// TwinCAT 3 PLC project PLC_Tank
// ProgramVersion: 3.1.4026.27
// libraries:
//   Tc2_ControllerToolbox, * (Beckhoff Automation GmbH)
//   Tc2_ModbusSrv, * (Beckhoff Automation GmbH)
//   Tc2_Standard, * (Beckhoff Automation GmbH)
//   Tc2_System, * (Beckhoff Automation GmbH)
//   Tc3_Module, * (Beckhoff Automation GmbH)
//   VisuDialogs, * (System)
//   VisuSymbols,3.5.10.0,System
// project tree:
//   DUTs/ TAnalogConversion.TcDUT, TEngine.TcDUT, TEngineCmd.TcDUT, THeaterState.TcDUT, THeaterCmd.TcDUT, THeater.TcDUT, TPhaseHeating.TcDUT, TPhaseCmd.TcDUT, TPhaseDraining.TcDUT, TPhaseFilling.TcDUT, TPhaseMixing.TcDUT, TPhaseState.TcDUT, TValveState.TcDUT, TValveCmd.TcDUT, TEngineState.TcDUT, TTank.TcDUT, TValve.TcDUT
//   / GlobalTextList.TcGTLO, PlcTask.TcTTO, PlcTask500ms.TcTTO, VisualizationManager.TcVMO (not stored)
//   GVLs/ Global.TcGVL
//   POUs/ Draining.TcPOU, Engine_1DO.TcPOU, FB_Tank.TcPOU, Filling.TcPOU, Heater.TcPOU, Heating.TcPOU, Main_Batch.TcPOU, MB_Connector.TcPOU, Mixing.TcPOU, Test.TcPOU, Valve_2DO.TcPOU, MAIN.TcPOU
//   POUs/Misc/ EngToRaw.TcPOU, RawToEng.TcPOU
//   VISUs/ Diagnostika.TcVIS, Faze.TcVIS, Prehled.TcVIS, Zarizeni.TcVIS
// real-time tasks:
//   TASK PlcTask: cycle T#100000us, priority 20, ADS port 350
//   TASK PlcTask500ms: cycle T#500ms, priority 1, ADS port 351

CONFIGURATION PLC_Tank
    RESOURCE PLC ON TwinCAT3
        TASK PlcTask(INTERVAL := T#100000us, PRIORITY := 20);
        TASK PlcTask500ms(INTERVAL := T#500ms, PRIORITY := 1);
        PROGRAM MB_Connector WITH PlcTask : MB_Connector;
        PROGRAM Main_Batch WITH PlcTask : Main_Batch;
        PROGRAM MAIN WITH PlcTask500ms : MAIN;
    END_RESOURCE
END_CONFIGURATION

// ---- DUTs/TAnalogConversion.TcDUT
TYPE TAnalogConversion :
STRUCT
	TransducerLoLevel : UINT;
	TransducerHiLevel : UINT;
	ScaledValLoLevel : REAL;
	ScaledValHiLevel : REAL;
END_STRUCT
END_TYPE

// ---- DUTs/TEngine.TcDUT
TYPE TEngine :
STRUCT
	Cmd : TEngineCmd;
	State : TEngineState;
	Time2Start : TIME := T#5S;
	RisingEdgeTrigger : R_TRIG;
	StartupFailTimer : TON;
END_STRUCT
END_TYPE

// ---- DUTs/TEngineCmd.TcDUT
TYPE TEngineCmd :
STRUCT
		SetRT : DINT;
		AutCtrl : BOOL;
		ManCtrl : BOOL;
		TurnOnMan : BOOL;
		TurnOffMan : BOOL;
		Req2RunAutCtrl : BOOL;
		ResetSUF : BOOL;
END_STRUCT
END_TYPE

// ---- DUTs/THeaterState.TcDUT
TYPE THeaterState :
STRUCT
	EnableOut : BOOL;
	HeatingOut : REAL;
	AutCtrl : BOOL;
	ManCtrl : BOOL;
	Err 	: BOOL;
	StateInt : INT;
	GenErr : BOOL; //signalisation: error occured

	HeatingPower : REAL;
	

END_STRUCT
END_TYPE

// ---- DUTs/THeaterCmd.TcDUT
TYPE THeaterCmd :
STRUCT
	AutCtrl : BOOL;
	ManCtrl : BOOL;
	TurnOnMan : BOOL;
	TurnOffMan : BOOL;
	Req2RunAutCtrl : BOOL;
END_STRUCT
END_TYPE

// ---- DUTs/THeater.TcDUT
TYPE THeater :
STRUCT
	Cmd : THeaterCmd;
	State : THeaterState;
	
	ParamHeatingPowerManual : REAL;
	ParamHeatingSetPointAutomat : REAL;
	
	PID : FB_CTRL_PID;
	ThresholdTimer : TON;
	
END_STRUCT
END_TYPE

// ---- DUTs/TPhaseHeating.TcDUT
TYPE TPhaseHeating :
STRUCT
	Cmd : TPhaseCmd;
	State : TPhaseState;
	
	ParamReqTemp : REAL;
	
	WaterTemp : REAL;
	
	fTime : INT;
END_STRUCT
END_TYPE

// ---- DUTs/TPhaseCmd.TcDUT
TYPE TPhaseCmd :
STRUCT
	StartAut : BOOL;
	StopAut : BOOL;
	StartMan : BOOL;
	StopMan : BOOL;
	PauseMan : BOOL;
	ResumeMan : BOOL;
	ResetDone : BOOL;
	AutCtrl : BOOL;
	ManCtrl : BOOL;
END_STRUCT
END_TYPE

// ---- DUTs/TPhaseDraining.TcDUT
TYPE TPhaseDraining :
STRUCT
	Cmd : TPhaseCmd;
	State : TPhaseState;
	
	ParamDrainLevel : REAL;
	WaterLevel : REAL;
END_STRUCT
END_TYPE

// ---- DUTs/TPhaseFilling.TcDUT
TYPE TPhaseFilling :
STRUCT
	Cmd : TPhaseCmd;
	State : TPhaseState;
	
	ParamFillLevel : REAL;
	WaterLevel : REAL;
END_STRUCT
END_TYPE

// ---- DUTs/TPhaseMixing.TcDUT
TYPE TPhaseMixing :
STRUCT
	Cmd : TPhaseCmd;
	State : TPhaseState;
	
	ParamTimeSec : INT;
	
	ElapsedTimeSec : INT;
END_STRUCT
END_TYPE

// ---- DUTs/TPhaseState.TcDUT
TYPE TPhaseState :
STRUCT
	Running : BOOL;
	Idle : BOOL;
	Paused : BOOL;
	Done : BOOL;
	AutCtrl : BOOL;
	ManCtrl : BOOL;
	Stateint : INT;
END_STRUCT
END_TYPE

// ---- DUTs/TValveState.TcDUT
TYPE TValveState :
STRUCT
		Open : BOOL;
		Closed : BOOL;
		OpenOut : BOOL;
		CloseOut : BOOL;
		Err : BOOL;
		StartupFail : BOOL;
		AutCtrl : BOOL;
		ManCtrl : BOOL;
		MayRun : BOOL;
		MayAutoRun : BOOL; //device is working in automatic regime
		GenErr : BOOL; //signalisation: error occured
		StColor : INT; //valve state: Open(0), Closed(1), OpenAndErr(2), ClosedAndErr(3) ,NotOpenNotClosedNotErr(4), NotOpenNotClosedAndErr(5), OpenAndClosedAndErr(6), OpenAndClosedNotErr(7)

END_STRUCT
END_TYPE

// ---- DUTs/TValveCmd.TcDUT
TYPE TValveCmd :
STRUCT
		AutCtrl : BOOL;
		ManCtrl : BOOL;
		OpenMan : BOOL;
		StopMan : BOOL;
		CloseMan : BOOL;
		Req2OpenAut : BOOL;
		Req2CloseAut : BOOL;
		ResetSUF : BOOL;
END_STRUCT
END_TYPE

// ---- DUTs/TEngineState.TcDUT
TYPE TEngineState :
STRUCT
		RT : DINT;
		Run : BOOL;
		RunOut : BOOL;
		Err : BOOL;
		StartUpFail : BOOL;
		AutCtrl : BOOL;
		ManCtrl : BOOL;
		MayRun : BOOL;
		MayAutoRun : BOOL;
		GenErr : BOOL;
		StateInt : INT;
		
		StartupFailTime : INT;
END_STRUCT
END_TYPE

// ---- DUTs/TTank.TcDUT
TYPE TTank :
STRUCT
	Mixer : TEngine;
	ValveFilling : TValve;
	ValveDraining : TValve;
	Heater : THeater;
	
	Filling : TPhaseFilling;
	Draining : TPhaseDraining;
	Mixing : TPhaseMixing;
	Heating : TPhaseHeating;
	
	GlobalError : BOOL;

END_STRUCT
END_TYPE

// ---- DUTs/TValve.TcDUT
TYPE TValve :
STRUCT
	Cmd : TValveCmd;
	State : TValveState;
	Time2Open : TIME := T#12S;
	
	OpenFailTimer : TON;
	CloseFailTimer : TON;
	
END_STRUCT
END_TYPE

// ---- GVLs/Global.TcGVL
{attribute 'qualified_only'}
VAR_GLOBAL
	Tank1 : TTank;
	

	secImp : BOOL;
	
	diMixerRun : BOOL;
	diMixerError : BOOL;
	diValveFillOpen : BOOL;
	diValveFillClose : BOOL;
	diValveFillError : BOOL;
	diValveDrainOpen : BOOL;
	diValveDrainClose : BOOL;
	diValveDrainError : BOOL;
	
	aiWaterLevel : WORD;
	aiWaterTemp : WORD;
	
	doMixerStart : BOOL;
	doValveFillOpen : BOOL;
	doValveFillClose : BOOL;
	doValveDrainOpen : BOOL;
	doValveDrainClose : BOOL;
	doHeatingEnable : BOOL;
	
	aoReqPowerOfHeating : WORD;

END_VAR

VAR_GLOBAL CONSTANT
	Running : INT := 0;
	Stop : INT := 1;
	RunningAndError : INT := 2;
	Err : INT := 3;

	PhIdle : INT := 0;
	PhRunning : INT := 1;
	PhPause : INT := 2;
	
    Open : INT := 0;
	Closed : INT := 1;
	OpenAndErr : INT := 2;
	ClosedAndErr : INT := 3;
	NotOpenNotClosedNotErr : INT := 4;
	NotOpenNotClosedAndErr : INT := 5;
	OpenAndClosedAndErr : INT := 6;
	OpenAndClosedNotErr : INT := 7;
END_VAR

// ---- POUs/MB_Connector.TcPOU
PROGRAM MB_Connector
VAR
	
	mb_ipaddr   : STRING(15) := '127.0.0.1';
	mb_port		: UINT := 504;
	mb_unitid	: BYTE := 1;
	
	fbReadRegs		: FB_MBReadInputRegs;
	mb_regs    		: ARRAY [0..4] OF WORD;
	mb_regs_error	: BOOL;
	mb_regs_busy	: BOOL;
	mb_regs_execute : BOOL;
	mb_regs_errid	: UDINT;
	
	fbReadInps	: FB_MBReadInputs;
	mb_inps			: ARRAY [0..4] OF BYTE;
	mb_inps_error	: BOOL;
	mb_inps_busy	: BOOL;
	mb_inps_execute : BOOL;
	mb_inps_errid	: UDINT;
	
	fbWriteRegs		: FB_MBWriteRegs;
	mbw_regs    	: ARRAY [0..4] OF WORD;
	mbw_regs_error	: BOOL;
	mbw_regs_busy	: BOOL;
	mbw_regs_execute: BOOL;
	mbw_regs_errid	: UDINT;
	
	fbWriteCoils	: FB_MBWriteCoils;
	mbw_coils		: ARRAY [0..4] OF BYTE;
	mbw_coils_error	: BOOL;
	mbw_coils_busy	: BOOL;
	mbw_coils_execute: BOOL;
	mbw_coils_errid	: UDINT;
	
END_VAR

fbReadRegs.sIPAddr := mb_ipaddr;
fbReadRegs.nTCPPort := mb_port;
fbReadRegs.nQuantity := 4;
fbReadRegs.nMBAddr := 0;
fbReadRegs.cbLength := SIZEOF(mb_regs);
fbReadRegs.pDestAddr := ADR(mb_regs);
fbReadRegs.nUnitID := mb_unitid;
fbReadRegs.tTimeout := T#5S;
IF (mb_regs_busy = FALSE) THEN
	mb_regs_execute := TRUE;
ELSE
	mb_regs_execute := FALSE;
END_IF
fbReadRegs(bExecute := mb_regs_execute, 
		   bBusy => mb_regs_busy, bError => mb_regs_error, 
		   nErrId => mb_regs_errid);



fbReadInps.sIPAddr := mb_ipaddr;
fbReadInps.nTCPPort := mb_port;
fbReadInps.nQuantity := 32;
fbReadInps.nMBAddr := 0;
fbReadInps.cbLength := SIZEOF(mb_inps);
fbReadInps.pDestAddr := ADR(mb_inps);
fbReadInps.nUnitID := mb_unitid;
fbReadInps.tTimeout := T#5S;
IF (mb_inps_busy = FALSE) THEN
	mb_inps_execute := TRUE;
ELSE
	mb_inps_execute := FALSE;
END_IF
fbReadInps(bExecute := mb_inps_execute, 
	bBusy => mb_inps_busy, bError => mb_inps_error, nErrId => mb_inps_errid);

Global.diValveFillOpen := mb_inps[0].0;
Global.diValveFillClose := mb_inps[0].1;
Global.diValveFillError := mb_inps[0].2;
Global.diValveDrainOpen := mb_inps[0].3;
Global.diValveDrainClose := mb_inps[0].4;
Global.diValveDrainError := mb_inps[0].5;
Global.diMixerRun := mb_inps[0].6;
Global.diMixerError := mb_inps[0].7;

Global.aiWaterLevel := mb_regs[0];
Global.aiWaterTemp := mb_regs[2];







fbWriteRegs.sIPAddr := mb_ipaddr;
fbWriteRegs.nTCPPort := mb_port;
fbWriteRegs.nQuantity := 4;
fbWriteRegs.nMBAddr := 0;
fbWriteRegs.cbLength := SIZEOF(mbw_regs);
fbWriteRegs.pSrcAddr := ADR(mbw_regs);
fbWriteRegs.nUnitID := mb_unitid;
fbWriteRegs.tTimeout := T#5S;
IF (mbw_regs_busy = FALSE) THEN
	mbw_regs_execute := TRUE;
ELSE
	mbw_regs_execute := FALSE;
END_IF
fbWriteRegs(bExecute := mbw_regs_execute, 
		   bBusy => mbw_regs_busy, bError => mbw_regs_error, 
		   nErrId => mbw_regs_errid);



fbWriteCoils.sIPAddr := mb_ipaddr;
fbWriteCoils.nTCPPort := mb_port;
fbWriteCoils.nQuantity := 32;
fbWriteCoils.nMBAddr := 0;
fbWriteCoils.cbLength := SIZEOF(mbw_coils);
fbWriteCoils.pSrcAddr := ADR(mbw_coils);
fbWriteCoils.nUnitID := mb_unitid;
fbWriteCoils.tTimeout := T#5S;
IF (mbw_coils_busy = FALSE) THEN
	mbw_coils_execute := TRUE;
ELSE
	mbw_coils_execute := FALSE;
END_IF
fbWriteCoils(bExecute := mbw_coils_execute, 
	bBusy => mbw_coils_busy, bError => mbw_coils_error, nErrId => mbw_coils_errid);

mbw_coils[0].0 := Global.doValveFillOpen;
mbw_coils[0].1 := Global.doValveFillClose;
mbw_coils[0].2 := Global.doValveDrainOpen;
mbw_coils[0].3 := Global.doValveDrainClose;
mbw_coils[0].4 := Global.doMixerStart;
mbw_coils[0].5 := Global.doHeatingEnable;

mbw_regs[0] := Global.aoReqPowerOfHeating;

END_PROGRAM

// ---- POUs/Main_Batch.TcPOU
PROGRAM Main_Batch
VAR
	FB_Tank_1 : FB_Tank;
END_VAR

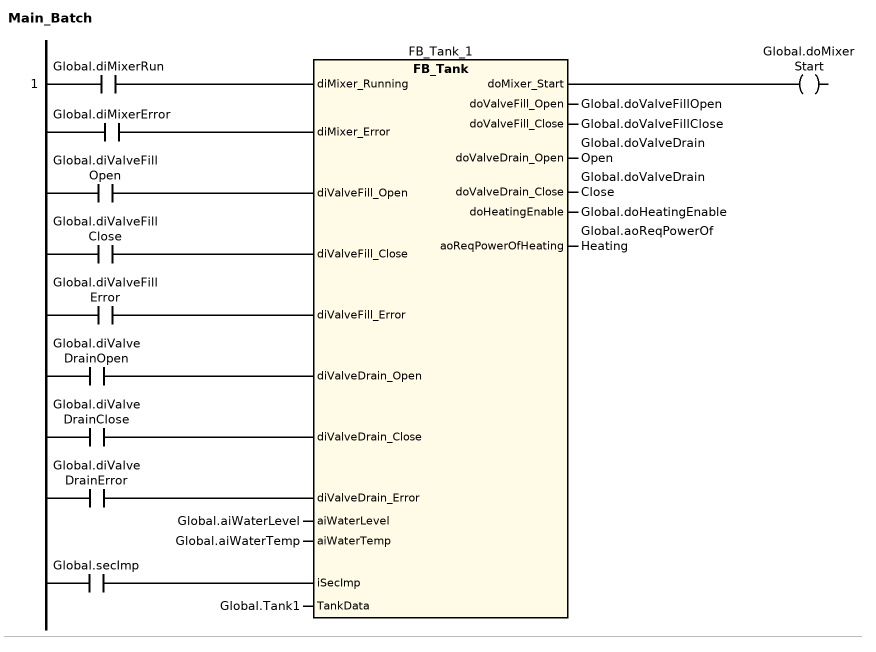
// NETWORK 1
FB_Tank_1(
    diMixer_Running := Global.diMixerRun,
    diMixer_Error := Global.diMixerError,
    diValveFill_Open := Global.diValveFillOpen,
    diValveFill_Close := Global.diValveFillClose,
    diValveFill_Error := Global.diValveFillError,
    diValveDrain_Open := Global.diValveDrainOpen,
    diValveDrain_Close := Global.diValveDrainClose,
    diValveDrain_Error := Global.diValveDrainError,
    aiWaterLevel := Global.aiWaterLevel,
    aiWaterTemp := Global.aiWaterTemp,
    iSecImp := Global.secImp,
    TankData := Global.Tank1,
    doValveFill_Open => Global.doValveFillOpen,
    doValveFill_Close => Global.doValveFillClose,
    doValveDrain_Open => Global.doValveDrainOpen,
    doValveDrain_Close => Global.doValveDrainClose,
    doHeatingEnable => Global.doHeatingEnable,
    aoReqPowerOfHeating => Global.aoReqPowerOfHeating); // FB_Tank
Global.doMixerStart := FB_Tank_1.doMixer_Start;

END_PROGRAM

// ---- POUs/FB_Tank.TcPOU
FUNCTION_BLOCK FB_Tank
VAR_INPUT
	diMixer_Running : BOOL;
	diMixer_Error : BOOL;
	diValveFill_Open : BOOL;
	diValveFill_Close : BOOL;
	diValveFill_Error : BOOL;
	diValveDrain_Open : BOOL;
	diValveDrain_Close : BOOL;
	diValveDrain_Error : BOOL;
	aiWaterLevel : WORD;
	aiWaterTemp : WORD;
	iSecImp : BOOL; //Požaduje se vstup s periodou 1 sekunda a libovolnou střídou
END_VAR

VAR_OUTPUT
	doMixer_Start : BOOL;
	doValveFill_Open : BOOL;
	doValveFill_Close : BOOL;
	doValveDrain_Open : BOOL;
	doValveDrain_Close : BOOL;
	doHeatingEnable : BOOL;
	aoReqPowerOfHeating : WORD;
END_VAR

VAR_IN_OUT
	TankData : TTank;
END_VAR

VAR
	//Konfigurace přepočtu rozsahu převodníků
	WaterTemp : TAnalogConversion := (TransducerLoLevel := 0, TransducerHiLevel := 27648, ScaledValLoLevel := 0, ScaledValHiLevel := 100);
	WaterLevel : TAnalogConversion := (TransducerLoLevel := 0, TransducerHiLevel := 27648, ScaledValLoLevel := 0, ScaledValHiLevel := 2);
	ReqOutputPower : TAnalogConversion := (ScaledValLoLevel := 0, ScaledValHiLevel := 100, TransducerLoLevel := 0, TransducerHiLevel := 27648);

	//Instance zanořených funkčních bloků
	ValveDrainCm : Valve_2DO;
	ValveFillCm : Valve_2DO;
	MixerCm : Engine_1DO;
	HeaterCm : Heater;
	FillingPhase : Filling;
	MixingPhase : Mixing;
	DrainingPhase : Draining;
	HeatingPhase : Heating;
	TON1: TON;
	RawToEng_1: RawToEng;
	RawToEng_2: RawToEng;
	EngToRaw_1: EngToRaw;
END_VAR

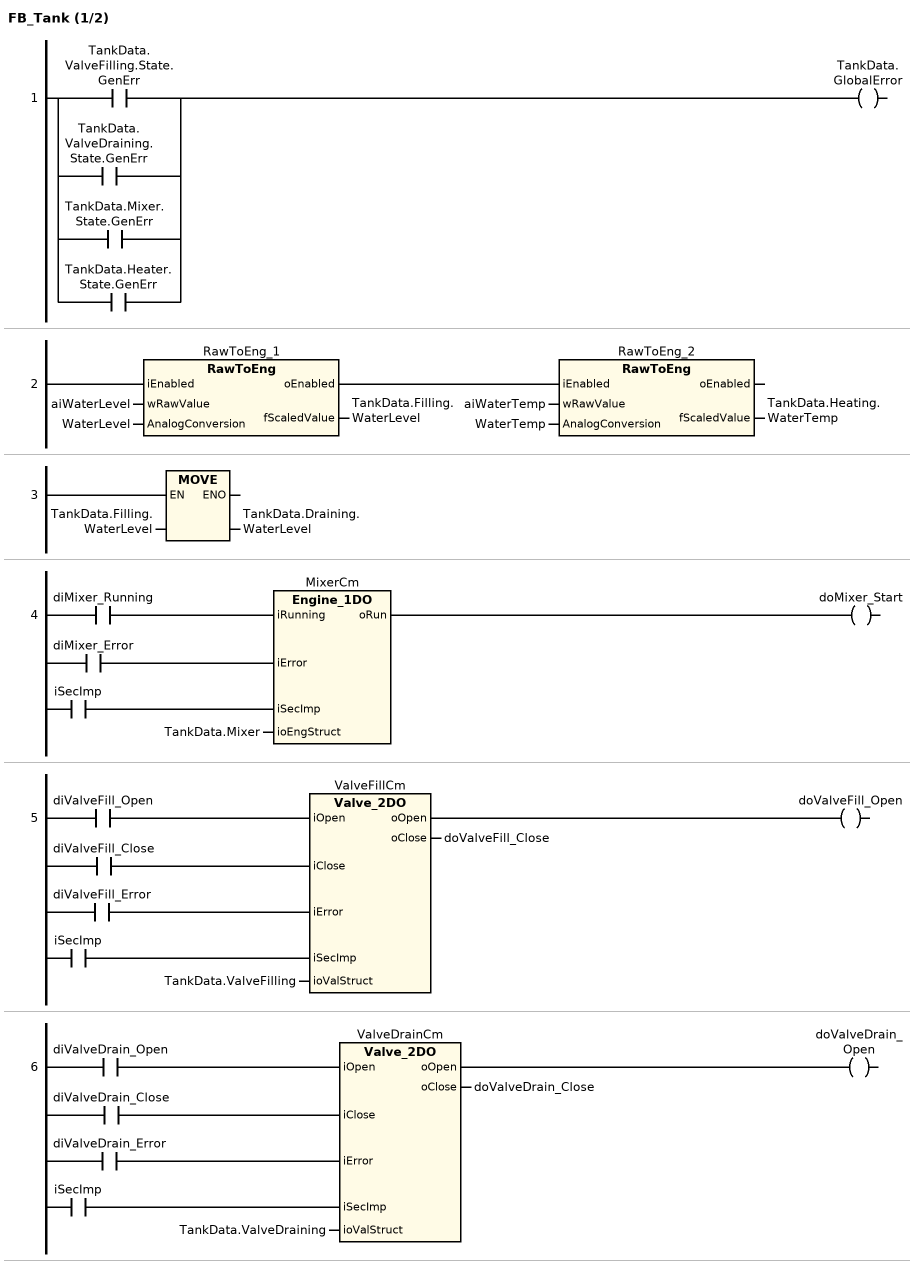
// NETWORK 1
TankData.GlobalError := TankData.ValveFilling.State.GenErr OR TankData.ValveDraining.State.GenErr OR TankData.Mixer.State.GenErr OR TankData.Heater.State.GenErr;

// NETWORK 2
RawToEng_1(
    iEnabled := TRUE,
    wRawValue := aiWaterLevel,
    AnalogConversion := WaterLevel,
    fScaledValue => TankData.Filling.WaterLevel); // RawToEng
RawToEng_2(
    iEnabled := RawToEng_1.oEnabled,
    wRawValue := aiWaterTemp,
    AnalogConversion := WaterTemp,
    fScaledValue => TankData.Heating.WaterTemp); // RawToEng

// NETWORK 3
TankData.Draining.WaterLevel := TankData.Filling.WaterLevel;

// NETWORK 4
MixerCm(
    iRunning := diMixer_Running,
    iError := diMixer_Error,
    iSecImp := iSecImp,
    ioEngStruct := TankData.Mixer); // Engine_1DO
doMixer_Start := MixerCm.oRun;

// NETWORK 5
ValveFillCm(
    iOpen := diValveFill_Open,
    iClose := diValveFill_Close,
    iError := diValveFill_Error,
    iSecImp := iSecImp,
    ioValStruct := TankData.ValveFilling,
    oClose => doValveFill_Close); // Valve_2DO
doValveFill_Open := ValveFillCm.oOpen;

// NETWORK 6
ValveDrainCm(
    iOpen := diValveDrain_Open,
    iClose := diValveDrain_Close,
    iError := diValveDrain_Error,
    iSecImp := iSecImp,
    ioValStruct := TankData.ValveDraining,
    oClose => doValveDrain_Close); // Valve_2DO
doValveDrain_Open := ValveDrainCm.oOpen;

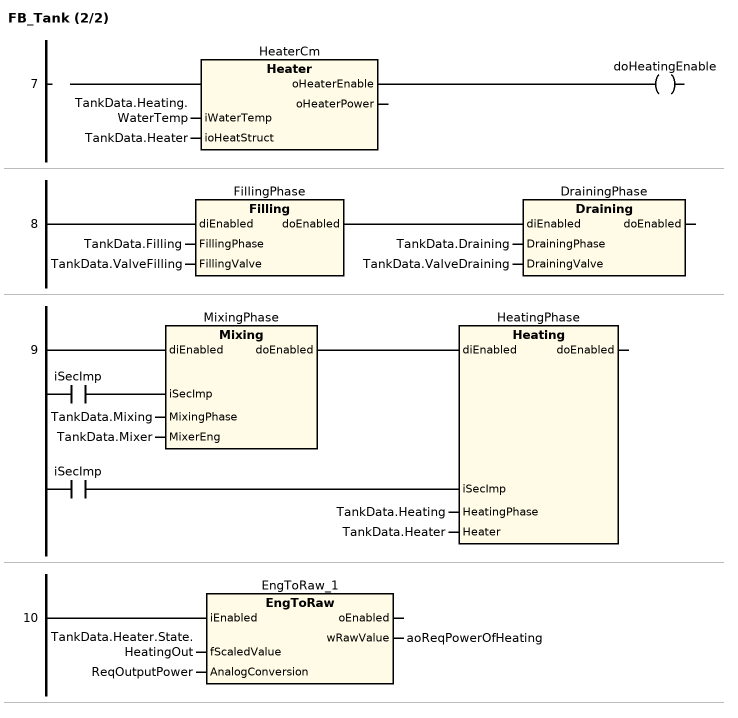
// NETWORK 7
HeaterCm(iWaterTemp := TankData.Heating.WaterTemp, ioHeatStruct := TankData.Heater); // Heater
doHeatingEnable := HeaterCm.oHeaterEnable;

// NETWORK 8
FillingPhase(diEnabled := TRUE, FillingPhase := TankData.Filling, FillingValve := TankData.ValveFilling); // Filling
DrainingPhase(
    diEnabled := FillingPhase.doEnabled,
    DrainingPhase := TankData.Draining,
    DrainingValve := TankData.ValveDraining); // Draining

// NETWORK 9
MixingPhase(
    diEnabled := TRUE,
    iSecImp := iSecImp,
    MixingPhase := TankData.Mixing,
    MixerEng := TankData.Mixer); // Mixing
HeatingPhase(
    diEnabled := MixingPhase.doEnabled,
    iSecImp := iSecImp,
    HeatingPhase := TankData.Heating,
    Heater := TankData.Heater); // Heating

// NETWORK 10
EngToRaw_1(
    iEnabled := TRUE,
    fScaledValue := TankData.Heater.State.HeatingOut,
    AnalogConversion := ReqOutputPower,
    wRawValue => aoReqPowerOfHeating); // EngToRaw

END_FUNCTION_BLOCK

// ---- POUs/Valve_2DO.TcPOU
FUNCTION_BLOCK Valve_2DO
VAR_INPUT
	iOpen : BOOL;
	iClose : BOOL;
	iError : BOOL;
	iSecImp : BOOL;
END_VAR
VAR_OUTPUT
	oOpen : BOOL;
	oClose : BOOL;
END_VAR

VAR_IN_OUT
	ioValStruct	 : TValve;
END_VAR

VAR
	tempOpenStartupFail : BOOL;
	tempCloseStartupFail: BOOL;
END_VAR

{region "OpenState"}
    // set real state of valve input into valve structure - input of valve can be taken from limit sensor...
    ioValStruct.State.Open := iOpen;
    ioValStruct.State.Closed := iClose;
{endregion}

	 
{region "REGION Aut/Man"}
    // switching state of engine - automatic or manual control (default state is manual)
  	IF ioValStruct.Cmd.ManCtrl THEN
      	ioValStruct.State.ManCtrl := TRUE;
		ioValStruct.State.AutCtrl := FALSE;
	ELSIF ioValStruct.Cmd.AutCtrl THEN
        ioValStruct.State.ManCtrl := FALSE;
		ioValStruct.State.AutCtrl := TRUE; 
    END_IF;
		 
	IF (NOT ioValStruct.State.AutCtrl AND NOT ioValStruct.State.ManCtrl) THEN
		ioValStruct.State.ManCtrl := TRUE;
	END_IF

	ioValStruct.Cmd.ManCtrl := FALSE;
	ioValStruct.Cmd.AutCtrl := FALSE;
{endregion}
	 
{region "MayRun / MayAutoRun"}
    // setting auxilary signals (may run, may auto run) - MR AND NOT MAR - engine may be started in manual mode, MAR - engine may be started in automatic mode
    ioValStruct.State.MayRun := (ioValStruct.State.ManCtrl AND NOT(ioValStruct.State.GenErr));
	ioValStruct.State.MayAutoRun := (ioValStruct.State.AutCtrl AND NOT(ioValStruct.State.GenErr));
{endregion}
	 
{region "ManCtrl"}
	// processing manual actions - if command is processed, it is sets to FALSE even if can't be processed
    // Valve commands are open, close and stop - valve can be stopped intermediate position
	 IF ioValStruct.State.ManCtrl AND ioValStruct.State.MayRun THEN
        IF ioValStruct.Cmd.OpenMan THEN
            ioValStruct.State.CloseOut := FALSE;
            ioValStruct.State.OpenOut := TRUE;
        END_IF;
        
        IF ioValStruct.Cmd.CloseMan THEN
            ioValStruct.State.OpenOut := FALSE;
            ioValStruct.State.CloseOut := TRUE;
        END_IF;
        
        IF ioValStruct.Cmd.StopMan THEN
            ioValStruct.State.OpenOut := FALSE;
            ioValStruct.State.CloseOut := FALSE;
        END_IF;
    END_IF;
    
    ioValStruct.Cmd.OpenMan := FALSE;
    ioValStruct.Cmd.CloseMan := FALSE;
    ioValStruct.Cmd.StopMan := FALSE;
{endregion}
	 
{region "AutCtrl"}
	 //if request to run in automatic mode -> set outputs to right states if MAR
    //AutoRequest shouldn't be reseted to false state
    //if request to open and request to close are setted to 1 simultaneously - outputs should be 0.
    IF ioValStruct.State.AutCtrl AND ioValStruct.State.MayAutoRun THEN
        IF ioValStruct.Cmd.Req2CloseAut AND (NOT ioValStruct.Cmd.Req2OpenAut) THEN
            ioValStruct.State.OpenOut := FALSE;
            ioValStruct.State.CloseOut := TRUE;
        END_IF;
        
        IF (NOT ioValStruct.Cmd.Req2CloseAut) AND ioValStruct.Cmd.Req2OpenAut THEN
            ioValStruct.State.CloseOut := FALSE;
            ioValStruct.State.OpenOut := TRUE;
        END_IF;
        
        IF (NOT ioValStruct.Cmd.Req2CloseAut) AND (NOT ioValStruct.Cmd.Req2OpenAut) THEN
            ioValStruct.State.CloseOut := FALSE;
            ioValStruct.State.OpenOut := FALSE;
        END_IF;
        
    END_IF;
{endregion}
	 
{region "Error states"}
 // definition of error states 
    // error - input from digital input of plc - fyzical state of valve
    // calculating start up fail - if output is sets to open or close, it's expected feedback from limit sensor in defined time, if feedback doesn't show in this time, it should be start up fail error
    // merge of these two error is general error
    // error is both inputs (open and closed) true state
    ioValStruct.OpenFailTimer(IN := ioValStruct.State.OpenOut AND NOT ioValStruct.State.CloseOut AND NOT ioValStruct.State.Open, PT := ioValStruct.Time2Open);
	tempOpenStartupFail := ioValStruct.OpenFailTimer.Q;

    ioValStruct.CloseFailTimer(IN := ioValStruct.State.CloseOut AND NOT ioValStruct.State.OpenOut AND NOT ioValStruct.State.Closed, PT := ioValStruct.Time2Open);
	tempCloseStartupFail := ioValStruct.CloseFailTimer.Q;
    
   
    IF tempOpenStartupFail OR tempCloseStartupFail THEN
        ioValStruct.State.StartUpFail := TRUE;
    END_IF;
    
    IF iError THEN
        ioValStruct.State.Err := TRUE;
    END_IF;
    
    ioValStruct.State.GenErr := ioValStruct.State.StartUpFail OR iError;
    
    // start up fail can be reseted by operator, command resetSUF, resets SUF and engine should be started again
    IF ioValStruct.Cmd.ResetSUF THEN
        ioValStruct.State.StartUpFail := FALSE;
        ioValStruct.Cmd.ResetSUF := FALSE;
    END_IF;
    
    // if error state exists outputs should be in stop state
    IF ioValStruct.State.GenErr THEN
        ioValStruct.State.OpenOut := FALSE;
        ioValStruct.State.CloseOut := FALSE;
    END_IF;
{endregion}
	 	 
oOpen := ioValStruct.State.OpenOut;
oClose := ioValStruct.State.CloseOut;

{region "StatusInt"}
    //write combination of states into int value for visualization (valve - combination of open, close state and error)
    IF ioValStruct.State.Open AND NOT ioValStruct.State.Closed AND NOT ioValStruct.State.GenErr THEN
        ioValStruct.State.StColor := Global.Open;
    ELSIF NOT ioValStruct.State.Open AND ioValStruct.State.Closed AND NOT ioValStruct.State.GenErr THEN
        ioValStruct.State.StColor := Global.Closed;
    ELSIF ioValStruct.State.Open AND NOT ioValStruct.State.Closed AND ioValStruct.State.GenErr THEN
        ioValStruct.State.StColor := Global.OpenAndErr;
    ELSIF NOT ioValStruct.State.Open AND ioValStruct.State.Closed AND ioValStruct.State.GenErr THEN
        ioValStruct.State.StColor := Global.ClosedAndErr;
    ELSIF NOT ioValStruct.State.Open AND NOT ioValStruct.State.Closed AND NOT ioValStruct.State.GenErr THEN
        ioValStruct.State.StColor := Global.NotOpenNotClosedNotErr;
    ELSIF NOT ioValStruct.State.Open AND NOT ioValStruct.State.Closed AND ioValStruct.State.GenErr THEN
        ioValStruct.State.StColor := Global.NotOpenNotClosedAndErr;
    ELSIF ioValStruct.State.Open AND ioValStruct.State.Closed AND ioValStruct.State.GenErr THEN
        ioValStruct.State.StColor := Global.OpenAndClosedAndErr;
    ELSIF ioValStruct.State.Open AND ioValStruct.State.Closed AND NOT ioValStruct.State.GenErr THEN
        ioValStruct.State.StColor := Global.OpenAndClosedNotErr;
    END_IF;
{endregion}

END_FUNCTION_BLOCK

// ---- POUs/Engine_1DO.TcPOU
FUNCTION_BLOCK Engine_1DO
VAR_INPUT
	iRunning : BOOL;
	iError : BOOL;
	iSecImp : BOOL;
END_VAR
VAR_OUTPUT
	oRun : BOOL;
END_VAR
VAR_IN_OUT
	ioEngStruct : TEngine;
END_VAR
VAR
	secImpEdge: BOOL;
	tempStartupFail: BOOL;
END_VAR

{region "RunState"}
    // set real state of engine run into engine structure
  ioEngStruct.State.Run := iRunning;
{endregion}

{region "Running time"} 
    // counting running time of engine - (motoseconds in real situation it should be moto hours)
    // detection rising edge of input secimp - should be conected 1Hz internal clock from PLC
	IF ioEngStruct.State.Run THEN
		IF iSecImp AND NOT secImpEdge THEN
			secImpEdge := TRUE;
			ioEngStruct.State.RT := ioEngStruct.State.RT + 1;
		ELSIF NOT iSecImp THEN
			secImpEdge := FALSE; 
		END_IF
	END_IF 
	
	IF ioEngStruct.Cmd.SetRT >= 0 THEN
		ioEngStruct.State.RT := ioEngStruct.Cmd.SetRT;
		ioEngStruct.Cmd.SetRT := -1;
	END_IF
{endregion}
	 
 
{region "Manual/Automat"}
	// switching state of engine - automatic or manual control (default state is manual)
	IF ioEngStruct.Cmd.ManCtrl THEN
      	ioEngStruct.State.ManCtrl := TRUE;
		ioEngStruct.State.AutCtrl := FALSE;
	ELSIF ioEngStruct.Cmd.AutCtrl THEN
        ioEngStruct.State.ManCtrl := FALSE;
		ioEngStruct.State.AutCtrl := TRUE; 
    END_IF;
		 
	IF (NOT ioEngStruct.State.AutCtrl AND NOT ioEngStruct.State.ManCtrl) THEN
		ioEngStruct.State.ManCtrl := TRUE;
	END_IF

	ioEngStruct.Cmd.ManCtrl := FALSE;
	ioEngStruct.Cmd.AutCtrl := FALSE;
{endregion}
	 
{region "MayRun / MayAutoRun"}
	// setting auxilary signals (may run, may auto run) - MR AND NOT MAR - eng should be started in manual mode,
    // MAR - should be started in automatic mode
    ioEngStruct.State.MayRun := (ioEngStruct.State.ManCtrl AND NOT(ioEngStruct.State.GenErr));
	ioEngStruct.State.MayAutoRun := (ioEngStruct.State.AutCtrl AND NOT(ioEngStruct.State.GenErr));  
{endregion}
	 
{region "ManCtrl"}
	// processing manual actions - if command is processed, it is set to FALSE even if can't be processed
    // Engine commands are turn off (stop) and turn on (start)
	IF ioEngStruct.State.ManCtrl AND ioEngStruct.State.MayRun THEN
		IF ioEngStruct.Cmd.TurnOnMan THEN
			ioEngStruct.State.RunOut := TRUE;
		ELSIF ioEngStruct.Cmd.TurnOffMan THEN
			ioEngStruct.State.RunOut := FALSE;
		END_IF
    END_IF;
	ioEngStruct.Cmd.TurnOnMan := FALSE;
	ioEngStruct.Cmd.TurnOffMan := FALSE;
{endregion}
	 
{region "AutCtrl"}
	//if request to run in automatic mode set outputs to right states if MAR
    //AutoRequest shouldn't be reseted to false state
    IF ioEngStruct.State.AutCtrl AND ioEngStruct.State.MayAutoRun THEN
		IF ioEngStruct.Cmd.Req2RunAutCtrl THEN
			ioEngStruct.State.RunOut := TRUE;
		ELSIF NOT ioEngStruct.Cmd.Req2RunAutCtrl THEN
			ioEngStruct.State.RunOut := FALSE;
		END_IF
    END_IF;
{endregion}
	 
{region "Error states"}
	// definition of error states 
	// error - input from digital input of plc - fyzical state of engine 
	// calculating start up fail - if output is sets to start engine, it's expected feedback from running signal in defined time, if feedback doesn't show in this time, it should be start up fail error
	// merge of these two error is general error
	ioEngStruct.StartupFailTimer(IN := ioEngStruct.State.RunOut AND NOT iRunning, PT := ioEngStruct.Time2Start);
    IF ioEngStruct.StartupFailTimer.Q THEN
        ioEngStruct.State.StartUpFail := TRUE;
    END_IF;

    ioEngStruct.State.Err := iError;
    ioEngStruct.State.GenErr := ioEngStruct.State.StartUpFail OR iError;

    IF ioEngStruct.Cmd.ResetSUF THEN
        ioEngStruct.State.StartUpFail := FALSE;
        ioEngStruct.Cmd.ResetSUF := FALSE;
    END_IF;

    IF ioEngStruct.State.GenErr THEN
        ioEngStruct.State.RunOut := FALSE;
    END_IF;
{endregion}
	 
oRun := ioEngStruct.State.RunOut;

{region "StatusInt"}
 IF NOT ioEngStruct.State.GenErr THEN
        IF ioEngStruct.State.Run THEN
            ioEngStruct.State.StateInt := Global.Running;
        ELSE
            ioEngStruct.State.StateInt := Global.Stop;
        END_IF;
    ELSE
        IF ioEngStruct.State.Run THEN
            ioEngStruct.State.StateInt := Global.RunningAndError;
        ELSE
            ioEngStruct.State.StateInt := Global.Err;
        END_IF;
    END_IF; 
{endregion}

END_FUNCTION_BLOCK

// ---- POUs/Heater.TcPOU
FUNCTION_BLOCK Heater
VAR_INPUT
	iWaterTemp : REAL;
END_VAR
VAR_OUTPUT
	oHeaterEnable : BOOL;
	oHeaterPower : REAL;
END_VAR
VAR_IN_OUT
	ioHeatStruct : THeater;
END_VAR
VAR
	pidParameters : ST_CTRL_PID_PARAMS;
	pidMode : E_CTRL_MODE;      // ACTIVE when heater is enabled, RESET otherwise
END_VAR

pidParameters.fKp := 1.196; //P
pidParameters.tTn := T#75.798S; //I
pidParameters.tTv := T#0S; //D
pidParameters.tCtrlCycleTime := T#200MS;
pidParameters.tTaskCycleTime := T#100MS;
pidParameters.fOutMaxLimit := 100;
pidParameters.fOutMinLimit := 0;
pidParameters.bDInTheFeedbackPath := FALSE;
pidParameters.bPInTheFeedbackPath := FALSE;
pidParameters.bARWOnIPartOnly := FALSE;
pidParameters.tTd := T#100MS; 


// PID runs only when heater is enabled - otherwise it is held in reset,
// so the integral part doesn't wind up while heating is off (no overshoot after start)
IF ioHeatStruct.State.EnableOut THEN
	pidMode := E_CTRL_MODE.eCTRL_MODE_ACTIVE;
ELSE
	pidMode := E_CTRL_MODE.eCTRL_MODE_RESET;
END_IF;

ioHeatStruct.PID(
	fSetpointValue := ioHeatStruct.ParamHeatingSetPointAutomat, 
	fActualValue := iWaterTemp, 
	fManSyncValue := ioHeatStruct.ParamHeatingPowerManual,
	bSync := ioHeatStruct.State.ManCtrl,
	eMode := pidMode, // automatic mode of PID component
	stParams := pidParameters);

ioHeatStruct.State.HeatingOut := ioHeatStruct.PID.fOut;

	 
{region "Manual/Automat"}
// switching state of engine - automatic or manual control (default state is manual)
	IF ioHeatStruct.Cmd.ManCtrl THEN
      	ioHeatStruct.State.ManCtrl := TRUE;
		ioHeatStruct.State.AutCtrl := FALSE;
	ELSIF ioHeatStruct.Cmd.AutCtrl THEN
        ioHeatStruct.State.ManCtrl := FALSE;
		ioHeatStruct.State.AutCtrl := TRUE; 
    END_IF;
		 
	IF (NOT ioHeatStruct.State.AutCtrl AND NOT ioHeatStruct.State.ManCtrl) THEN
		ioHeatStruct.State.ManCtrl := TRUE;
	END_IF

	ioHeatStruct.Cmd.ManCtrl := FALSE;
	ioHeatStruct.Cmd.AutCtrl := FALSE;
{endregion}
	 
 
{region "ManCtrl"}
	// processing manual actions - if command is processed, it is set to FALSE even if can't be processed
	// Heater commands are turn off (stop) and turn on (start) and power level
	IF ioHeatStruct.State.ManCtrl THEN
		IF ioHeatStruct.Cmd.TurnOnMan AND NOT ioHeatStruct.State.GenErr THEN
			ioHeatStruct.State.EnableOut := TRUE;
		ELSIF ioHeatStruct.Cmd.TurnOffMan THEN
			ioHeatStruct.State.EnableOut := FALSE;
		END_IF
    END_IF;
	ioHeatStruct.Cmd.TurnOnMan := FALSE;
	ioHeatStruct.Cmd.TurnOffMan := FALSE;
{endregion}
 
{region "AutCtrl"}
	//if request to run in automatic mode set outputs to right states if MAR
	//AutoRequest shouldn't be reseted to false state
    IF ioHeatStruct.State.AutCtrl THEN
		IF ioHeatStruct.Cmd.Req2RunAutCtrl AND NOT ioHeatStruct.State.GenErr THEN
			ioHeatStruct.State.EnableOut := TRUE;
		ELSIF NOT ioHeatStruct.Cmd.Req2RunAutCtrl THEN
			ioHeatStruct.State.EnableOut := FALSE;
		END_IF
    END_IF;
{endregion}
 
{region "Error states"}
	// if water temperature is too high, stop heating and generate error
	IF iWaterTemp > 90 THEN
		ioHeatStruct.State.EnableOut := FALSE;
		ioHeatStruct.State.GenErr := TRUE;
	ELSIF iWaterTemp < 85 THEN
		ioHeatStruct.State.GenErr := FALSE;
	END_IF
	ioHeatStruct.State.Err := ioHeatStruct.State.GenErr;
{endregion}
	 
 IF NOT ioHeatStruct.State.EnableOut THEN
    ioHeatStruct.State.HeatingOut := 0;
ELSIF ioHeatStruct.State.ManCtrl THEN
    ioHeatStruct.State.HeatingOut := ioHeatStruct.ParamHeatingPowerManual;
ELSE
    ioHeatStruct.State.HeatingOut := ioHeatStruct.PID.fOut;
END_IF;
 
oHeaterPower := ioHeatStruct.State.HeatingOut;
oHeaterEnable := ioHeatStruct.State.EnableOut;

END_FUNCTION_BLOCK

// ---- POUs/Filling.TcPOU
FUNCTION_BLOCK Filling
VAR_INPUT
	diEnabled : BOOL;
END_VAR
VAR_OUTPUT
	doEnabled : BOOL;
END_VAR
VAR_IN_OUT
	FillingPhase : TPhaseFilling;
	FillingValve : TValve;
END_VAR
VAR
END_VAR

{region "REGION Aut/Man"}
    // switching state of engine - automatic or manual control (default state is manual)
  	IF FillingPhase.Cmd.ManCtrl THEN
      	FillingPhase.State.ManCtrl := TRUE;
		FillingPhase.State.AutCtrl := FALSE;
	ELSIF FillingPhase.Cmd.AutCtrl THEN
        FillingPhase.State.ManCtrl := FALSE;
		FillingPhase.State.AutCtrl := TRUE; 
    END_IF;
		 
	IF (NOT FillingPhase.State.AutCtrl AND NOT FillingPhase.State.ManCtrl) THEN
		FillingPhase.State.ManCtrl := TRUE;
	END_IF

	FillingPhase.Cmd.ManCtrl := FALSE;
	FillingPhase.Cmd.AutCtrl := FALSE;
{endregion}

{region "ManCtrl"}
    // processing manual actions - if command is processed, it is sets to FALSE even if can't be processed
    // Phase commands are start, stop, pause and resume 
    // Start - open filling valve 
    // Stop - close filling valve
    // Pause - close filling valve
    // Resume - open filling valve
    // real states of phase are wrote into states in phase structure
    IF FillingPhase.State.ManCtrl THEN
		IF FillingPhase.State.Idle AND FillingPhase.Cmd.StartMan THEN
			FillingPhase.State.Running := TRUE;
			FillingPhase.State.Idle := FALSE;
			FillingPhase.State.Paused := FALSE;
		 	FillingPhase.State.Done := FALSE;
		ELSIF FillingPhase.Cmd.StopMan THEN
			FillingPhase.State.Running := FALSE;
			FillingPhase.State.Idle := TRUE;
			FillingPhase.State.Paused := FALSE;
		ELSIF FillingPhase.State.Running AND FillingPhase.Cmd.PauseMan THEN
			FillingPhase.State.Running := FALSE;
			FillingPhase.State.Idle := FALSE;
			FillingPhase.State.Paused := TRUE;
		ELSIF FillingPhase.State.Paused AND FillingPhase.Cmd.ResumeMan THEN
			FillingPhase.State.Running := TRUE;
			FillingPhase.State.Idle := FALSE;
			FillingPhase.State.Paused := FALSE;
			FillingPhase.State.Done := FALSE;
		END_IF
    END_IF;
	
	FillingPhase.Cmd.StartMan := FALSE;
	FillingPhase.Cmd.StopMan := FALSE;
	FillingPhase.Cmd.PauseMan := FALSE;
	FillingPhase.Cmd.ResumeMan := FALSE;
{endregion}

{region "AutCtrl"}
    // if request to run in automatic mode and phase can be run in automatic mode switch phase to running
    IF FillingPhase.State.AutCtrl THEN
		IF FillingPhase.State.Idle AND FillingPhase.Cmd.StartAut THEN
			FillingPhase.State.Running := TRUE;
			FillingPhase.State.Idle := FALSE;
		 	FillingPhase.State.Done := FALSE;
		ELSIF FillingPhase.Cmd.StopAut THEN
			FillingPhase.State.Running := FALSE;
			FillingPhase.State.Idle := TRUE;
			FillingPhase.State.Paused := FALSE;
		END_IF
    END_IF;
	
	FillingPhase.Cmd.StartAut := FALSE;
	FillingPhase.Cmd.StopAut := FALSE;
{endregion}

{region "Done"}
    //every phase should have finish condition - filling phase - if water level is above requested level
    //after that done state should be set to 1
    IF FillingPhase.State.Running AND (FillingPhase.WaterLevel >= FillingPhase.ParamFillLevel - 0.083) THEN // edit based on speed of simulation 
        FillingPhase.Cmd.StopMan := TRUE;
        FillingPhase.Cmd.StopAut := TRUE;
        FillingPhase.State.Done := TRUE;
    END_IF;

    IF FillingPhase.Cmd.ResetDone THEN
        FillingPhase.State.Done := FALSE;
        FillingPhase.Cmd.ResetDone := FALSE;
    END_IF;
{endregion}

{region "States"}
	//Command valve in cases of states
    IF FillingPhase.State.Running THEN
        FillingValve.Cmd.Req2OpenAut := TRUE;
        FillingValve.Cmd.Req2CloseAut := FALSE;
    ELSE
        FillingValve.Cmd.Req2OpenAut := FALSE;
        FillingValve.Cmd.Req2CloseAut := TRUE;
    END_IF;
{endregion}


// delault state of phase - if not any state sets state to idle
IF NOT FillingPhase.State.Idle AND NOT FillingPhase.State.Paused AND NOT FillingPhase.State.Running THEN
    FillingPhase.State.Idle := 1;
END_IF;

// write binary states into int value for visualization
IF FillingPhase.State.Idle THEN
    FillingPhase.State.Stateint := Global.PhIdle;
ELSIF FillingPhase.State.Running THEN
    FillingPhase.State.Stateint := Global.PhRunning;
ELSE
    FillingPhase.State.Stateint := Global.PhPause;
END_IF;

// Ponechte pro moznost retezeni volani bloku v LAD
doEnabled := diEnabled;

END_FUNCTION_BLOCK

// ---- POUs/Mixing.TcPOU
FUNCTION_BLOCK Mixing
VAR_INPUT
	diEnabled : BOOL;
	iSecImp : BOOL;
END_VAR
VAR_OUTPUT
	doEnabled : BOOL;
END_VAR
VAR_IN_OUT
	MixingPhase : TPhaseMixing;
	MixerEng : TEngine;
END_VAR
VAR
	rtSecImp : R_TRIG;          // rising edge of second impulse
END_VAR

{region "Aut/Man"}
    // switching state of phase - automatic or manual control (default state is manual)
    // if both commands come at once, manual has priority (safety)
    IF MixingPhase.Cmd.ManCtrl THEN
        MixingPhase.State.ManCtrl := TRUE;
        MixingPhase.State.AutCtrl := FALSE;
    ELSIF MixingPhase.Cmd.AutCtrl THEN
        MixingPhase.State.ManCtrl := FALSE;
        MixingPhase.State.AutCtrl := TRUE;
    END_IF;

    // initialization - if neither mode is active, use manual
    IF NOT MixingPhase.State.AutCtrl AND NOT MixingPhase.State.ManCtrl THEN
        MixingPhase.State.ManCtrl := TRUE;
    END_IF;

    // commands are always reset after processing
    MixingPhase.Cmd.ManCtrl := FALSE;
    MixingPhase.Cmd.AutCtrl := FALSE;
{endregion}

{region "ManCtrl"}
    // processing manual actions - if command is processed, it is set to FALSE even if can't be processed
    // Phase commands are start, stop, pause and resume
    // Start  - start mixing (elapsed time starts from 0)
    // Stop   - stop mixing
    // Pause  - stop mixing (elapsed time is kept)
    // Resume - start mixing (continues for the remaining time)
    IF MixingPhase.State.ManCtrl THEN
        IF MixingPhase.State.Idle AND MixingPhase.Cmd.StartMan THEN
            MixingPhase.State.Running := TRUE;
            MixingPhase.State.Idle := FALSE;
            MixingPhase.State.Paused := FALSE;
            MixingPhase.State.Done := FALSE;
            MixingPhase.ElapsedTimeSec := 0;
        ELSIF MixingPhase.Cmd.StopMan THEN
            MixingPhase.State.Running := FALSE;
            MixingPhase.State.Idle := TRUE;
            MixingPhase.State.Paused := FALSE;
        ELSIF MixingPhase.State.Running AND MixingPhase.Cmd.PauseMan THEN
            MixingPhase.State.Running := FALSE;
            MixingPhase.State.Idle := FALSE;
            MixingPhase.State.Paused := TRUE;
        ELSIF MixingPhase.State.Paused AND MixingPhase.Cmd.ResumeMan THEN
            MixingPhase.State.Running := TRUE;
            MixingPhase.State.Idle := FALSE;
            MixingPhase.State.Paused := FALSE;
            MixingPhase.State.Done := FALSE;
        END_IF;
    END_IF;

    MixingPhase.Cmd.StartMan := FALSE;
    MixingPhase.Cmd.StopMan := FALSE;
    MixingPhase.Cmd.PauseMan := FALSE;
    MixingPhase.Cmd.ResumeMan := FALSE;
{endregion}

{region "AutCtrl"}
    // if phase is in automatic mode, process StartAut / StopAut (from MES)
    // commands are set to FALSE after their processing
    IF MixingPhase.State.AutCtrl THEN
        IF MixingPhase.State.Idle AND MixingPhase.Cmd.StartAut THEN
            MixingPhase.State.Running := TRUE;
            MixingPhase.State.Idle := FALSE;
            MixingPhase.State.Done := FALSE;
            MixingPhase.ElapsedTimeSec := 0;
        ELSIF MixingPhase.Cmd.StopAut THEN
            MixingPhase.State.Running := FALSE;
            MixingPhase.State.Idle := TRUE;
            MixingPhase.State.Paused := FALSE;
        END_IF;
    END_IF;

    MixingPhase.Cmd.StartAut := FALSE;
    MixingPhase.Cmd.StopAut := FALSE;
{endregion}

{region "Done"}
    // every phase should have finish condition - mixing phase - elapsed running time >= requested time
    // elapsed time is counted only while running (second impulse rising edge),
    // it is kept during pause and reset only on start
    rtSecImp(CLK := iSecImp);   // must be called every cycle, otherwise edges are lost

    IF MixingPhase.State.Running AND rtSecImp.Q THEN
        MixingPhase.ElapsedTimeSec := MixingPhase.ElapsedTimeSec + 1;
    END_IF;

    // finish condition met -> stop phase (processed next cycle) and signal Done
    IF MixingPhase.State.Running AND (MixingPhase.ElapsedTimeSec >= MixingPhase.ParamTimeSec) THEN
        MixingPhase.Cmd.StopMan := TRUE;
        MixingPhase.Cmd.StopAut := TRUE;
        MixingPhase.State.Done := TRUE;
    END_IF;

    // command reset done resets done state and then resets command
    IF MixingPhase.Cmd.ResetDone THEN
        MixingPhase.State.Done := FALSE;
        MixingPhase.Cmd.ResetDone := FALSE;
    END_IF;
{endregion}

{region "States"}
    // Command mixer in cases of states
    // Running - mixer runs
    // Idle    - mixer stopped
    // Paused  - mixer stopped
    IF MixingPhase.State.Running THEN
        MixerEng.Cmd.Req2RunAutCtrl := TRUE;
    ELSE
        MixerEng.Cmd.Req2RunAutCtrl := FALSE;
    END_IF;
{endregion}

// default state of phase - if not any state sets state to idle
IF NOT MixingPhase.State.Idle AND NOT MixingPhase.State.Paused AND NOT MixingPhase.State.Running THEN
    MixingPhase.State.Idle := 1;
END_IF;

// write binary states into int value for visualization
IF MixingPhase.State.Idle THEN
    MixingPhase.State.Stateint := Global.PhIdle;
ELSIF MixingPhase.State.Running THEN
    MixingPhase.State.Stateint := Global.PhRunning;
ELSE
    MixingPhase.State.Stateint := Global.PhPause;
END_IF;

doEnabled := diEnabled;

END_FUNCTION_BLOCK

// ---- POUs/Draining.TcPOU
FUNCTION_BLOCK Draining
VAR_INPUT
	diEnabled : BOOL;
END_VAR
VAR_OUTPUT
	doEnabled : BOOL;
END_VAR
VAR_IN_OUT
	DrainingPhase : TPhaseDraining;
	DrainingValve : TValve;
END_VAR
VAR
END_VAR

{region "Aut/Man"}
    // switching state of engine - automatic or manual control (default state is manual)
  	IF DrainingPhase.Cmd.ManCtrl THEN
      	DrainingPhase.State.ManCtrl := TRUE;
		DrainingPhase.State.AutCtrl := FALSE;
	ELSIF DrainingPhase.Cmd.AutCtrl THEN
        DrainingPhase.State.ManCtrl := FALSE;
		DrainingPhase.State.AutCtrl := TRUE; 
    END_IF;
		 
	IF (NOT DrainingPhase.State.AutCtrl AND NOT DrainingPhase.State.ManCtrl) THEN
		DrainingPhase.State.ManCtrl := TRUE;
	END_IF

	DrainingPhase.Cmd.ManCtrl := FALSE;
	DrainingPhase.Cmd.AutCtrl := FALSE;
{endregion}

{region "ManCtrl"}
    // processing manual actions - if command is processed, it is sets to FALSE even if can't be processed
    // Phase commands are start, stop, pause and resume 
    // Start - open draining valve 
    // Stop - close draining valve
    // Pause - close draining valve
    // Resume - open draining valve
    // real states of phase are writed into states in phase structure
    IF DrainingPhase.State.ManCtrl THEN
		IF DrainingPhase.State.Idle AND DrainingPhase.Cmd.StartMan THEN
			DrainingPhase.State.Running := TRUE;
			DrainingPhase.State.Idle := FALSE;
			DrainingPhase.State.Paused := FALSE;
		 	DrainingPhase.State.Done := FALSE;
		ELSIF DrainingPhase.Cmd.StopMan THEN
			DrainingPhase.State.Running := FALSE;
			DrainingPhase.State.Idle := TRUE;
			DrainingPhase.State.Paused := FALSE;
		ELSIF DrainingPhase.State.Running AND DrainingPhase.Cmd.PauseMan THEN
			DrainingPhase.State.Running := FALSE;
			DrainingPhase.State.Idle := FALSE;
			DrainingPhase.State.Paused := TRUE;
		ELSIF DrainingPhase.State.Paused AND DrainingPhase.Cmd.ResumeMan THEN
			DrainingPhase.State.Running := TRUE;
			DrainingPhase.State.Idle := FALSE;
			DrainingPhase.State.Paused := FALSE;
			DrainingPhase.State.Done := FALSE;
		END_IF
    END_IF;
	
	DrainingPhase.Cmd.StartMan := FALSE;
	DrainingPhase.Cmd.StopMan := FALSE;
	DrainingPhase.Cmd.PauseMan := FALSE;
	DrainingPhase.Cmd.ResumeMan := FALSE;
{endregion}

{region "AutCtrl"}
    //if request to run in automatic mode -> set auto request to open of filling valve to 1 and close to 0, if not open 0 close 1
    // commands should be sets to false after their processing
    IF DrainingPhase.State.AutCtrl THEN
		IF DrainingPhase.State.Idle AND DrainingPhase.Cmd.StartAut THEN
			DrainingPhase.State.Running := TRUE;
			DrainingPhase.State.Idle := FALSE;
		 	DrainingPhase.State.Done := FALSE;
		ELSIF DrainingPhase.Cmd.StopAut THEN
			DrainingPhase.State.Running := FALSE;
			DrainingPhase.State.Idle := TRUE;
			DrainingPhase.State.Paused := FALSE;
		END_IF
    END_IF;
	
	DrainingPhase.Cmd.StartAut := FALSE;
	DrainingPhase.Cmd.StopAut := FALSE;
{endregion}
{region "Done"}
    //every phase should have finish condition - draining phase - if water level is below requested level
    //after that done state should be setted to 1
    IF DrainingPhase.State.Running AND (DrainingPhase.WaterLevel <= DrainingPhase.ParamDrainLevel) THEN // edit based on speed of simulation 
        DrainingPhase.Cmd.StopMan := TRUE;
        DrainingPhase.Cmd.StopAut := TRUE;
        DrainingPhase.State.Done := TRUE;
    END_IF;

    IF DrainingPhase.Cmd.ResetDone THEN
        DrainingPhase.State.Done := FALSE;
        DrainingPhase.Cmd.ResetDone := FALSE;
    END_IF;
{endregion}

{region "States"} 
    //Command valve in cases of states
    IF DrainingPhase.State.Running THEN
        DrainingValve.Cmd.Req2OpenAut := TRUE;
        DrainingValve.Cmd.Req2CloseAut := FALSE;
    ELSE
        DrainingValve.Cmd.Req2OpenAut := FALSE;
        DrainingValve.Cmd.Req2CloseAut := TRUE;
    END_IF;
{endregion}

// delault state of phase - if not any state sets state to idle
IF (NOT DrainingPhase.State.Idle) AND (NOT DrainingPhase.State.Paused) AND (NOT DrainingPhase.State.Running) THEN
    DrainingPhase.State.Idle := 1;
END_IF;

// write binary states into int value for visualization
IF DrainingPhase.State.Idle THEN
    DrainingPhase.State.StateInt := Global.PhIdle;
ELSIF DrainingPhase.State.Running THEN
    DrainingPhase.State.StateInt := Global.PhRunning;
ELSE
    DrainingPhase.State.StateInt := Global.PhPause;
END_IF;

//Ponechte pro moznost retezeni volani bloku v LAD
doEnabled := diEnabled;

END_FUNCTION_BLOCK

// ---- POUs/Heating.TcPOU
FUNCTION_BLOCK Heating
VAR_INPUT
	diEnabled : BOOL;
	iSecImp : BOOL;
END_VAR
VAR_OUTPUT
	doEnabled : BOOL;
END_VAR
VAR_IN_OUT
	HeatingPhase : TPhaseHeating;
	Heater : THeater;
END_VAR
VAR
	//pidParameters : ST_CTRL_PID_PARAMS;   // unused - PID is in Heater
	rtSecImp : R_TRIG;          // rising edge of second impulse
END_VAR

{region "Aut/Man"}
    // switching state of phase - automatic or manual control (default state is manual)
    // if both commands come at once, manual has priority (safety)
    IF HeatingPhase.Cmd.ManCtrl THEN
        HeatingPhase.State.ManCtrl := TRUE;
        HeatingPhase.State.AutCtrl := FALSE;
    ELSIF HeatingPhase.Cmd.AutCtrl THEN
        HeatingPhase.State.ManCtrl := FALSE;
        HeatingPhase.State.AutCtrl := TRUE;
    END_IF;

    // initialization - if neither mode is active, use manual
    IF NOT HeatingPhase.State.AutCtrl AND NOT HeatingPhase.State.ManCtrl THEN
        HeatingPhase.State.ManCtrl := TRUE;
    END_IF;

    // commands are always reset after processing
    HeatingPhase.Cmd.ManCtrl := FALSE;
    HeatingPhase.Cmd.AutCtrl := FALSE;
{endregion}

{region "ManCtrl"}
    // processing manual actions - if command is processed, it is set to FALSE even if can't be processed
    // Phase commands are start, stop, pause and resume
    // Start  - start heating
    // Stop   - stop heating
    // Pause  - stop heating (remaining condition is evaluated again after resume)
    // Resume - start heating
    // real states of phase are written into states in phase structure
    IF HeatingPhase.State.ManCtrl THEN
        IF HeatingPhase.State.Idle AND HeatingPhase.Cmd.StartMan THEN
            HeatingPhase.State.Running := TRUE;
            HeatingPhase.State.Idle := FALSE;
            HeatingPhase.State.Paused := FALSE;
            HeatingPhase.State.Done := FALSE;
        ELSIF HeatingPhase.Cmd.StopMan THEN
            HeatingPhase.State.Running := FALSE;
            HeatingPhase.State.Idle := TRUE;
            HeatingPhase.State.Paused := FALSE;
        ELSIF HeatingPhase.State.Running AND HeatingPhase.Cmd.PauseMan THEN
            HeatingPhase.State.Running := FALSE;
            HeatingPhase.State.Idle := FALSE;
            HeatingPhase.State.Paused := TRUE;
        ELSIF HeatingPhase.State.Paused AND HeatingPhase.Cmd.ResumeMan THEN
            HeatingPhase.State.Running := TRUE;
            HeatingPhase.State.Idle := FALSE;
            HeatingPhase.State.Paused := FALSE;
            HeatingPhase.State.Done := FALSE;
        END_IF;
    END_IF;

    HeatingPhase.Cmd.StartMan := FALSE;
    HeatingPhase.Cmd.StopMan := FALSE;
    HeatingPhase.Cmd.PauseMan := FALSE;
    HeatingPhase.Cmd.ResumeMan := FALSE;
{endregion}

{region "AutCtrl"}
    // if phase is in automatic mode, process StartAut / StopAut (from MES)
    // commands are set to FALSE after their processing
    IF HeatingPhase.State.AutCtrl THEN
        IF HeatingPhase.State.Idle AND HeatingPhase.Cmd.StartAut THEN
            HeatingPhase.State.Running := TRUE;
            HeatingPhase.State.Idle := FALSE;
            HeatingPhase.State.Done := FALSE;
        ELSIF HeatingPhase.Cmd.StopAut THEN
            HeatingPhase.State.Running := FALSE;
            HeatingPhase.State.Idle := TRUE;
            HeatingPhase.State.Paused := FALSE;
        END_IF;
    END_IF;

    HeatingPhase.Cmd.StartAut := FALSE;
    HeatingPhase.Cmd.StopAut := FALSE;
{endregion}

{region "Done"}
    // every phase should have finish condition - heating phase - water temp must stay
    // within +-1 °C of requested value for 10 seconds (skripta 10.3.11)
    // fTime counts seconds in tolerance band; it is reset when temp leaves the band or phase is not running
    rtSecImp(CLK := iSecImp);   // must be called every cycle, otherwise edges are lost

    IF HeatingPhase.State.Running THEN
        IF ABS(HeatingPhase.WaterTemp - HeatingPhase.ParamReqTemp) <= 1.0 THEN
            IF rtSecImp.Q THEN
                HeatingPhase.fTime := HeatingPhase.fTime + 1;
            END_IF;
        ELSE
            HeatingPhase.fTime := 0;
        END_IF;
    ELSE
        HeatingPhase.fTime := 0;
    END_IF;

    // finish condition met -> stop phase (processed next cycle) and signal Done
    IF HeatingPhase.State.Running AND (HeatingPhase.fTime >= 10) THEN
        HeatingPhase.Cmd.StopMan := TRUE;
        HeatingPhase.Cmd.StopAut := TRUE;
        HeatingPhase.State.Done := TRUE;
    END_IF;

    // command reset done resets done state and then resets command
    IF HeatingPhase.Cmd.ResetDone THEN
        HeatingPhase.State.Done := FALSE;
        HeatingPhase.Cmd.ResetDone := FALSE;
    END_IF;
{endregion}

{region "States"}
    // Command heater in cases of states
    // Running - start heating, pass requested temperature to heater (PID setpoint)
    // Idle    - stop heating
    // Paused  - stop heating (alternative would be holding actual temperature)
    IF HeatingPhase.State.Running THEN
        Heater.ParamHeatingSetPointAutomat := HeatingPhase.ParamReqTemp;
        Heater.Cmd.Req2RunAutCtrl := TRUE;
    ELSE
        Heater.Cmd.Req2RunAutCtrl := FALSE;
    END_IF;
{endregion}

// default state of phase - if not any state sets state to idle
IF NOT HeatingPhase.State.Idle AND NOT HeatingPhase.State.Paused AND NOT HeatingPhase.State.Running THEN
    HeatingPhase.State.Idle := 1;
END_IF;

// write binary states into int value for visualization
IF HeatingPhase.State.Idle THEN
    HeatingPhase.State.Stateint := Global.PhIdle;
ELSIF HeatingPhase.State.Running THEN
    HeatingPhase.State.Stateint := Global.PhRunning;
ELSE
    HeatingPhase.State.Stateint := Global.PhPause;
END_IF;

doEnabled := diEnabled;

END_FUNCTION_BLOCK

// ---- POUs/Misc/RawToEng.TcPOU
FUNCTION_BLOCK RawToEng
VAR_INPUT
	iEnabled : BOOL;
	wRawValue : WORD;
	AnalogConversion : TAnalogConversion;
END_VAR
VAR_OUTPUT
	oEnabled : BOOL;
	fScaledValue : REAL;
END_VAR
VAR
END_VAR

//Prepocet z wRawValue (z procesu po ModbusTCP) na fScaledValue (do PLC) podle parametru v AnalogConversion.

//Filtrace hodnoty, bylo by vhodne odfiltrovat take kmitani z minimalniho rozsahu na maximalni hodnotu 27648
IF wRawValue = 27648 THEN 
	wRawValue := 0; //Ale lepe nez takto...
END_IF

fScaledValue:= (AnalogConversion.ScaledValHiLevel-AnalogConversion.ScaledValLoLevel) * (wRawValue-AnalogConversion.TransducerLoLevel)/(AnalogConversion.TransducerHiLevel-AnalogConversion.TransducerLoLevel) + AnalogConversion.ScaledValLoLevel;
oEnabled := iEnabled;

END_FUNCTION_BLOCK

// ---- POUs/Misc/EngToRaw.TcPOU
FUNCTION_BLOCK EngToRaw
VAR_INPUT
	iEnabled : BOOL;
	fScaledValue : REAL;
	AnalogConversion : TAnalogConversion;
END_VAR
VAR_OUTPUT
	oEnabled : BOOL;
	wRawValue : WORD;
END_VAR
VAR
END_VAR

//Prepocet z fScaledValue (z PLC) na wRawValue (do procesu po ModbusTCP) podle parametru v AnalogConversion.
wRawValue := REAL_TO_WORD((AnalogConversion.TransducerHiLevel - AnalogConversion.TransducerLoLevel) * (fScaledValue - AnalogConversion.ScaledValLoLevel) / (AnalogConversion.ScaledValHiLevel - AnalogConversion.ScaledValLoLevel) + AnalogConversion.TransducerLoLevel);
oEnabled := iEnabled;

END_FUNCTION_BLOCK

// ---- POUs/MAIN.TcPOU
PROGRAM MAIN
VAR

END_VAR

Global.secImp := NOT(Global.secImp);

END_PROGRAM

// ---- POUs/Test.TcPOU
PROGRAM Test
VAR
	State : INT := 0;
END_VAR

CASE State OF
	1:  Global.Tank1.Filling.ParamFillLevel := 1.8;
		Global.Tank1.Filling.Cmd.ManCtrl := TRUE;
		Global.Tank1.Filling.Cmd.StartMan:= TRUE;
		IF Global.Tank1.Filling.State.Done = TRUE THEN
			State := 2;
		END_IF
	2: //...
END_CASE

END_PROGRAM

// ---- GlobalTextList.TcGTLO
TEXTLIST GlobalTextList
  1001 = 'Přehled'
  1002 = 'Manuál'
  1003 = 'Automat'
  1004 = 'Diagnostika'
  1005 = '%.2f m'
  1006 = '%.1f °C'
  1007 = 'GlobalError'
  1008 = 'V-plnění'
  1009 = 'V-vypouštění'
  1010 = 'Míchadlo'
  1011 = 'Ohřev'
  1012 = 'Hodnoty'
  1013 = 'Hladina'
  1014 = 'Teplota'
  1015 = 'Výkon ohřevu [%]'
  1016 = '%.1f %%'
  1017 = 'Zařízení'
  1018 = 'běží / otevř.'
  1019 = 'Fáze'
  1020 = 'Idle'
  1021 = 'Running'
  1022 = 'Paused'
  1023 = 'Done'
  1024 = 'Napouštění'
  1025 = 'Míchání'
  1026 = 'Vypouštění'
  1027 = 'Napouštěcí ventil'
  1028 = 'Otevřeno'
  1029 = 'Zavřeno'
  1030 = 'Porucha'
  1031 = 'Stop'
  1032 = 'Reset SUF'
  1033 = 'Běží'
  1034 = 'Zapnout'
  1035 = 'Vypnout'
  1036 = 'Motohodiny'
  1037 = '%d s'
  1038 = 'Vypouštěcí ventil'
  1039 = 'Zapnuto'
  1040 = '> 95 °C'
  1041 = 'Výkon manuál [%]'
  1042 = 'Nádrž'
  1043 = 'FillLevel [m]'
  1044 = '%.2f'
  1045 = 'Start'
  1046 = 'Pause'
  1047 = 'Resume'
  1048 = 'Reset Done'
  1049 = 'Doba míchání [s]'
  1050 = '%d'
  1051 = 'Uběhlo [s]'
  1052 = 'Teplota [°C]'
  1053 = 'Stabilní [s]'
  1054 = 'DrainLevel [m]'
  1055 = 'AUT = fázi řídí MES / recept v PLC, MAN = obsluha tlačítky na této stránce.'
  1056 = 'Modbus TCP'
  1057 = 'IP adresa'
  1058 = '%s'
  1059 = 'Port'
  1060 = 'Busy'
  1061 = 'Error'
  1062 = 'Error ID'
  1063 = 'Čtení registrů (0x04)'
  1064 = 'Čtení vstupů (0x02)'
  1065 = 'Zápis registrů (0x10)'
  1066 = 'Zápis cívek (0x0F)'
  1067 = 'Poruchy'
  1068 = 'StartupFail'
  1069 = 'StartUpFail'
  1070 = 'Porucha měniče'
  1071 = 'Přehřátí > 95 °C'
  1072 = 'Motohodiny [s]'
  1073 = 'Nastavit motohodiny [s]'
  994 = '%.1f'
  815 = 'ABC'
  406 = 'AUT'
  473 = 'Checkbox'
  70 = 'Close'
  25 = 'Closed'
  201 = 'Filling Valve'
  560 = 'MAN'
  604 = 'Open'
  687 = 'Opened'
  98 = 'Res. SUF'
  256 = 'SUF'
END_TEXTLIST

// ---- VISUs/Diagnostika.TcVIS
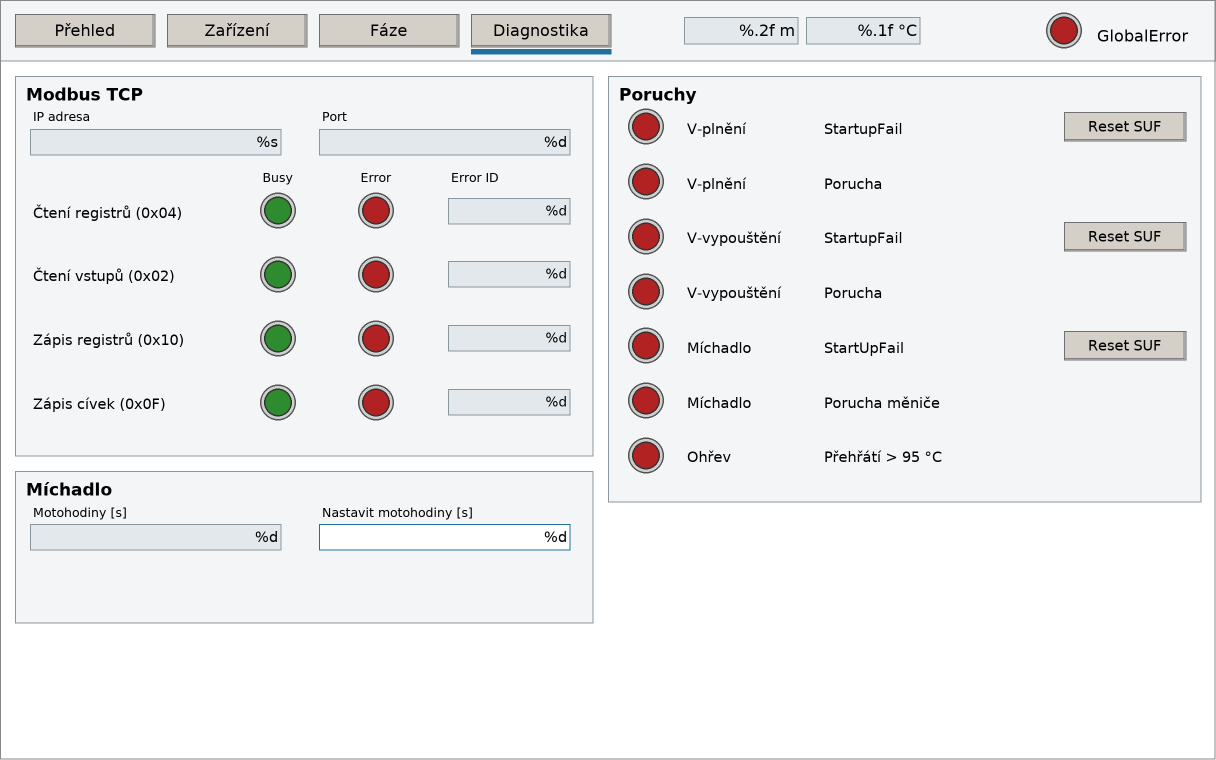
VISUALIZATION Diagnostika  // 1216x760
    Rectangle (0,0 1216x61)
    Button (15,14 140x33), "Přehled"
        OnMouseClick: change screen: Prehled
    Button (167,14 140x33), "Zařízení"
        OnMouseClick: change screen: Zarizeni
    Button (319,14 140x33), "Fáze"
        OnMouseClick: change screen: Faze
    Button (471,14 140x33), "Diagnostika"
        OnMouseClick: change screen: Diagnostika
    Rectangle (471,49 140x5)
    Rectangle (684,17 114x27), "%.2f m", text variable: Global.Tank1.Filling.WaterLevel
    Rectangle (806,17 114x27), "%.1f °C", text variable: Global.Tank1.Heating.WaterTemp
    Lamp1 (1041,10 46x41), variable: Global.Tank1.GlobalError, style: Lamp-Lamp1-Red
    Label (1094,23 126x26), "GlobalError"
    Rectangle (15,76 578x380)
    Label (23,81 122x27), "Modbus TCP"
    Label (30,106 83x21), "IP adresa"
    Rectangle (30,129 251x26), "%s", text variable: MB_Connector.mb_ipaddr
    Label (319,106 41x21), "Port"
    Rectangle (319,129 251x26), "%d", text variable: MB_Connector.mb_port
    Label (236,167 84x21), "Busy"
    Label (334,167 84x21), "Error"
    Label (433,167 84x21), "Error ID"
    Label (30,201 209x24), "Čtení registrů (0x04)"
    Lamp1 (255,190 46x41), variable: MB_Connector.mb_regs_busy, style: Lamp-Lamp1-Green
    Lamp1 (353,190 46x41), variable: MB_Connector.mb_regs_error, style: Lamp-Lamp1-Red
    Rectangle (448,198 122x26), "%d", text variable: MB_Connector.mb_regs_errid
    Label (30,264 190x24), "Čtení vstupů (0x02)"
    Lamp1 (255,254 46x41), variable: MB_Connector.mb_inps_busy, style: Lamp-Lamp1-Green
    Lamp1 (353,254 46x41), variable: MB_Connector.mb_inps_error, style: Lamp-Lamp1-Red
    Rectangle (448,261 122x26), "%d", text variable: MB_Connector.mb_inps_errid
    Label (30,328 209x24), "Zápis registrů (0x10)"
    Lamp1 (255,318 46x41), variable: MB_Connector.mbw_regs_busy, style: Lamp-Lamp1-Green
    Lamp1 (353,318 46x41), variable: MB_Connector.mbw_regs_error, style: Lamp-Lamp1-Red
    Rectangle (448,325 122x26), "%d", text variable: MB_Connector.mbw_regs_errid
    Label (30,392 180x24), "Zápis cívek (0x0F)"
    Lamp1 (255,382 46x41), variable: MB_Connector.mbw_coils_busy, style: Lamp-Lamp1-Green
    Lamp1 (353,382 46x41), variable: MB_Connector.mbw_coils_error, style: Lamp-Lamp1-Red
    Rectangle (448,389 122x26), "%d", text variable: MB_Connector.mbw_coils_errid
    Rectangle (608,76 593x426)
    Label (616,81 87x27), "Poruchy"
    Lamp1 (623,106 46x41), variable: Global.Tank1.ValveFilling.State.StartupFail, style: Lamp-Lamp1-Red
    Label (684,117 84x24), "V-plnění"
    Label (821,117 113x24), "StartupFail"
    Button (1064,112 122x29), "Reset SUF", colour toggle: Global.Tank1.ValveFilling.State.StartupFail
        tap Global.Tank1.ValveFilling.Cmd.ResetSUF
    Lamp1 (623,161 46x41), variable: Global.Tank1.ValveFilling.State.Err, style: Lamp-Lamp1-Red
    Label (684,172 84x24), "V-plnění"
    Label (821,172 74x24), "Porucha"
    Lamp1 (623,216 46x41), variable: Global.Tank1.ValveDraining.State.StartupFail, style: Lamp-Lamp1-Red
    Label (684,226 123x24), "V-vypouštění"
    Label (821,226 113x24), "StartupFail"
    Button (1064,222 122x29), "Reset SUF", colour toggle: Global.Tank1.ValveDraining.State.StartupFail
        tap Global.Tank1.ValveDraining.Cmd.ResetSUF
    Lamp1 (623,271 46x41), variable: Global.Tank1.ValveDraining.State.Err, style: Lamp-Lamp1-Red
    Label (684,281 123x24), "V-vypouštění"
    Label (821,281 74x24), "Porucha"
    Lamp1 (623,325 46x41), variable: Global.Tank1.Mixer.State.StartUpFail, style: Lamp-Lamp1-Red
    Label (684,336 84x24), "Míchadlo"
    Label (821,336 113x24), "StartUpFail"
    Button (1064,331 122x29), "Reset SUF", colour toggle: Global.Tank1.Mixer.State.StartUpFail
        tap Global.Tank1.Mixer.Cmd.ResetSUF
    Lamp1 (623,380 46x41), variable: Global.Tank1.Mixer.State.Err, style: Lamp-Lamp1-Red
    Label (684,391 84x24), "Míchadlo"
    Label (821,391 142x24), "Porucha měniče"
    Lamp1 (623,435 46x41), variable: Global.Tank1.Heater.State.GenErr, style: Lamp-Lamp1-Red
    Label (684,445 55x24), "Ohřev"
    Label (821,445 161x24), "Přehřátí > 95 °C"
    Rectangle (15,471 578x152)
    Label (23,476 99x27), "Míchadlo"
    Label (30,502 125x21), "Motohodiny [s]"
    Rectangle (30,524 251x26), "%d", text variable: Global.Tank1.Mixer.State.RT
    Label (319,502 201x21), "Nastavit motohodiny [s]"
    Rectangle (319,524 251x26), "%d", text variable: Global.Tank1.Mixer.Cmd.SetRT
        OnMouseClick: write the text variable via Default
END_VISUALIZATION

// ---- VISUs/Faze.TcVIS
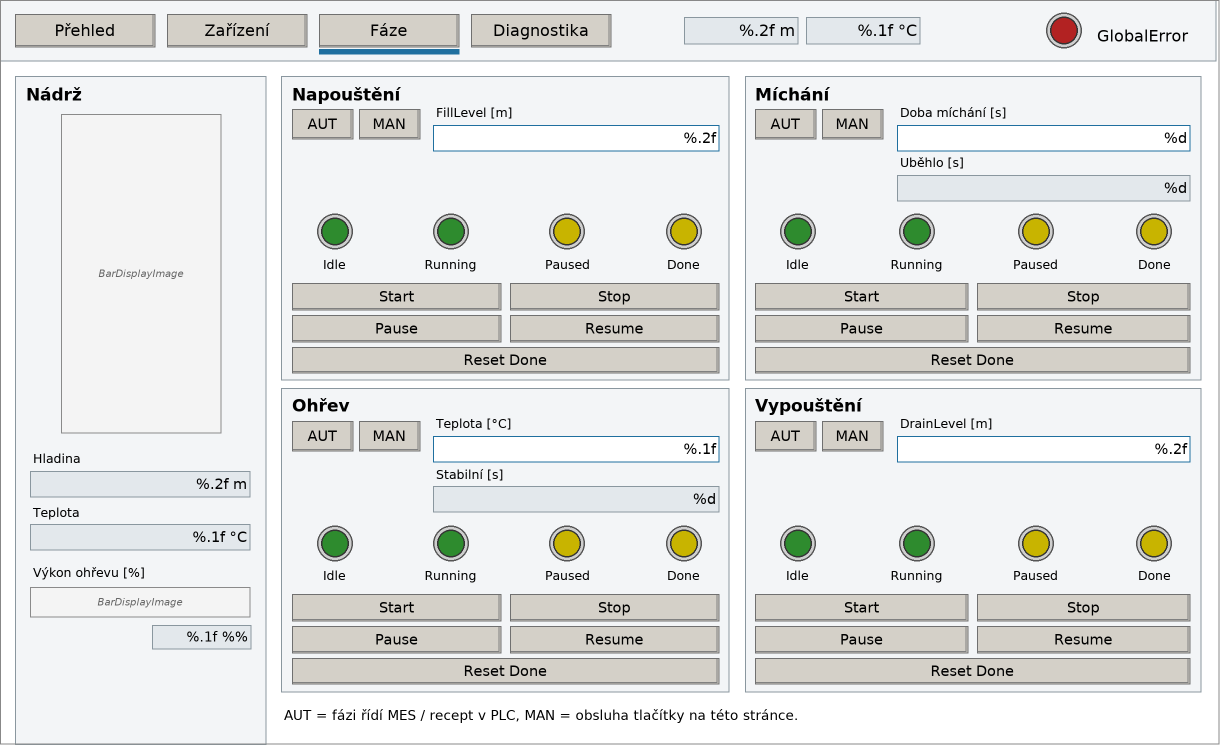
VISUALIZATION Faze  // 1220x745
    Rectangle (0,0 1216x61)
    Button (15,14 140x33), "Přehled"
        OnMouseClick: change screen: Prehled
    Button (167,14 140x33), "Zařízení"
        OnMouseClick: change screen: Zarizeni
    Button (319,14 140x33), "Fáze"
        OnMouseClick: change screen: Faze
    Rectangle (319,49 140x5)
    Button (471,14 140x33), "Diagnostika"
        OnMouseClick: change screen: Diagnostika
    Rectangle (684,17 114x27), "%.2f m", text variable: Global.Tank1.Filling.WaterLevel
    Rectangle (806,17 114x27), "%.1f °C", text variable: Global.Tank1.Heating.WaterTemp
    Lamp1 (1041,10 46x41), variable: Global.Tank1.GlobalError, style: Lamp-Lamp1-Red
    Label (1094,23 126x26), "GlobalError"
    Rectangle (15,76 251x669)
    Label (23,81 65x27), "Nádrž"
    BarDisplayImage (61,114 160x319), value: Global.Tank1.Filling.WaterLevel, style: BarDisplayImage-Gray, scale format: %.1f, scale 0..2
    Label (30,448 66x21), "Hladina"
    Rectangle (30,471 220x26), "%.2f m", text variable: Global.Tank1.Filling.WaterLevel
    Label (30,502 66x21), "Teplota"
    Rectangle (30,524 220x26), "%.1f °C", text variable: Global.Tank1.Heating.WaterTemp
    Label (30,562 142x21), "Výkon ohřevu [%]"
    BarDisplayImage (30,587 220x30), value: Global.Tank1.Heater.State.HeatingOut, style: BarDisplayImage-Gray, scale format: %.1f, scale 0..100
    Rectangle (152,625 99x24), "%.1f %%", text variable: Global.Tank1.Heater.State.HeatingOut
    Rectangle (281,76 448x304)
    Label (289,81 122x27), "Napouštění"
    Button (292,109 61x30), "AUT", colour toggle: Global.Tank1.Filling.State.AutCtrl
        tap Global.Tank1.Filling.Cmd.AutCtrl
    Button (359,109 61x30), "MAN", colour toggle: Global.Tank1.Filling.State.ManCtrl
        tap Global.Tank1.Filling.Cmd.ManCtrl
    Label (433,102 117x21), "FillLevel [m]"
    Rectangle (433,125 286x26), "%.2f", text variable: Global.Tank1.Filling.ParamFillLevel
        OnMouseClick: write the text variable via Default
    Lamp1 (312,211 46x41), variable: Global.Tank1.Filling.State.Idle, style: Lamp-Lamp1-Green
    Label (289,254 91x21), "Idle"
    Lamp1 (428,211 46x41), variable: Global.Tank1.Filling.State.Running, style: Lamp-Lamp1-Green
    Label (405,254 91x21), "Running"
    Lamp1 (544,211 46x41), variable: Global.Tank1.Filling.State.Paused, style: Lamp-Lamp1-Yellow
    Label (522,254 91x21), "Paused"
    Lamp1 (661,211 46x41), variable: Global.Tank1.Filling.State.Done, style: Lamp-Lamp1-Yellow
    Label (638,254 91x21), "Done"
    Button (292,283 209x27), "Start", colour toggle: Global.Tank1.Filling.State.Running
        tap Global.Tank1.Filling.Cmd.StartMan
    Button (510,283 209x27), "Stop"
        tap Global.Tank1.Filling.Cmd.StopMan
    Button (292,315 209x27), "Pause", colour toggle: Global.Tank1.Filling.State.Paused
        tap Global.Tank1.Filling.Cmd.PauseMan
    Button (510,315 209x27), "Resume"
        tap Global.Tank1.Filling.Cmd.ResumeMan
    Button (292,347 427x26), "Reset Done", colour toggle: Global.Tank1.Filling.State.Done
        tap Global.Tank1.Filling.Cmd.ResetDone
    Rectangle (745,76 456x304)
    Label (752,81 87x27), "Míchání"
    Button (755,109 61x30), "AUT", colour toggle: Global.Tank1.Mixing.State.AutCtrl
        tap Global.Tank1.Mixing.Cmd.AutCtrl
    Button (822,109 61x30), "MAN", colour toggle: Global.Tank1.Mixing.State.ManCtrl
        tap Global.Tank1.Mixing.Cmd.ManCtrl
    Label (897,102 142x21), "Doba míchání [s]"
    Rectangle (897,125 293x26), "%d", text variable: Global.Tank1.Mixing.ParamTimeSec
        OnMouseClick: write the text variable via Default
    Label (897,152 92x21), "Uběhlo [s]"
    Rectangle (897,175 293x26), "%d", text variable: Global.Tank1.Mixing.ElapsedTimeSec
    Lamp1 (775,211 46x41), variable: Global.Tank1.Mixing.State.Idle, style: Lamp-Lamp1-Green
    Label (752,254 91x21), "Idle"
    Lamp1 (894,211 46x41), variable: Global.Tank1.Mixing.State.Running, style: Lamp-Lamp1-Green
    Label (871,254 91x21), "Running"
    Lamp1 (1013,211 46x41), variable: Global.Tank1.Mixing.State.Paused, style: Lamp-Lamp1-Yellow
    Label (990,254 91x21), "Paused"
    Lamp1 (1131,211 46x41), variable: Global.Tank1.Mixing.State.Done, style: Lamp-Lamp1-Yellow
    Label (1109,254 91x21), "Done"
    Button (755,283 213x27), "Start", colour toggle: Global.Tank1.Mixing.State.Running
        tap Global.Tank1.Mixing.Cmd.StartMan
    Button (977,283 213x27), "Stop"
        tap Global.Tank1.Mixing.Cmd.StopMan
    Button (755,315 213x27), "Pause", colour toggle: Global.Tank1.Mixing.State.Paused
        tap Global.Tank1.Mixing.Cmd.PauseMan
    Button (977,315 213x27), "Resume"
        tap Global.Tank1.Mixing.Cmd.ResumeMan
    Button (755,347 435x26), "Reset Done", colour toggle: Global.Tank1.Mixing.State.Done
        tap Global.Tank1.Mixing.Cmd.ResetDone
    Rectangle (281,388 448x304)
    Label (289,392 65x27), "Ohřev"
    Button (292,421 61x30), "AUT", colour toggle: Global.Tank1.Heating.State.AutCtrl
        tap Global.Tank1.Heating.Cmd.AutCtrl
    Button (359,421 61x30), "MAN", colour toggle: Global.Tank1.Heating.State.ManCtrl
        tap Global.Tank1.Heating.Cmd.ManCtrl
    Label (433,413 109x21), "Teplota [°C]"
    Rectangle (433,436 286x26), "%.1f", text variable: Global.Tank1.Heating.ParamReqTemp
        OnMouseClick: write the text variable via Default
    Label (433,464 109x21), "Stabilní [s]"
    Rectangle (433,486 286x26), "%d", text variable: Global.Tank1.Heating.fTime
    Lamp1 (312,523 46x41), variable: Global.Tank1.Heating.State.Idle, style: Lamp-Lamp1-Green
    Label (289,565 91x21), "Idle"
    Lamp1 (428,523 46x41), variable: Global.Tank1.Heating.State.Running, style: Lamp-Lamp1-Green
    Label (405,565 91x21), "Running"
    Lamp1 (544,523 46x41), variable: Global.Tank1.Heating.State.Paused, style: Lamp-Lamp1-Yellow
    Label (522,565 91x21), "Paused"
    Lamp1 (661,523 46x41), variable: Global.Tank1.Heating.State.Done, style: Lamp-Lamp1-Yellow
    Label (638,565 91x21), "Done"
    Button (292,594 209x27), "Start", colour toggle: Global.Tank1.Heating.State.Running
        tap Global.Tank1.Heating.Cmd.StartMan
    Button (510,594 209x27), "Stop"
        tap Global.Tank1.Heating.Cmd.StopMan
    Button (292,626 209x27), "Pause", colour toggle: Global.Tank1.Heating.State.Paused
        tap Global.Tank1.Heating.Cmd.PauseMan
    Button (510,626 209x27), "Resume"
        tap Global.Tank1.Heating.Cmd.ResumeMan
    Button (292,658 427x26), "Reset Done", colour toggle: Global.Tank1.Heating.State.Done
        tap Global.Tank1.Heating.Cmd.ResetDone
    Rectangle (745,388 456x304)
    Label (752,392 122x27), "Vypouštění"
    Button (755,421 61x30), "AUT", colour toggle: Global.Tank1.Draining.State.AutCtrl
        tap Global.Tank1.Draining.Cmd.AutCtrl
    Button (822,421 61x30), "MAN", colour toggle: Global.Tank1.Draining.State.ManCtrl
        tap Global.Tank1.Draining.Cmd.ManCtrl
    Label (897,413 125x21), "DrainLevel [m]"
    Rectangle (897,436 293x26), "%.2f", text variable: Global.Tank1.Draining.ParamDrainLevel
        OnMouseClick: write the text variable via Default
    Lamp1 (775,523 46x41), variable: Global.Tank1.Draining.State.Idle, style: Lamp-Lamp1-Green
    Label (752,565 91x21), "Idle"
    Lamp1 (894,523 46x41), variable: Global.Tank1.Draining.State.Running, style: Lamp-Lamp1-Green
    Label (871,565 91x21), "Running"
    Lamp1 (1013,523 46x41), variable: Global.Tank1.Draining.State.Paused, style: Lamp-Lamp1-Yellow
    Label (990,565 91x21), "Paused"
    Lamp1 (1131,523 46x41), variable: Global.Tank1.Draining.State.Done, style: Lamp-Lamp1-Yellow
    Label (1109,565 91x21), "Done"
    Button (755,594 213x27), "Start", colour toggle: Global.Tank1.Draining.State.Running
        tap Global.Tank1.Draining.Cmd.StartMan
    Button (977,594 213x27), "Stop"
        tap Global.Tank1.Draining.Cmd.StopMan
    Button (755,626 213x27), "Pause", colour toggle: Global.Tank1.Draining.State.Paused
        tap Global.Tank1.Draining.Cmd.PauseMan
    Button (977,626 213x27), "Resume"
        tap Global.Tank1.Draining.Cmd.ResumeMan
    Button (755,658 435x26), "Reset Done", colour toggle: Global.Tank1.Draining.State.Done
        tap Global.Tank1.Draining.Cmd.ResetDone
    Label (281,704 682x23), "AUT = fázi řídí MES / recept v PLC, MAN = obsluha tlačítky na této stránce."
END_VISUALIZATION

// ---- VISUs/Prehled.TcVIS
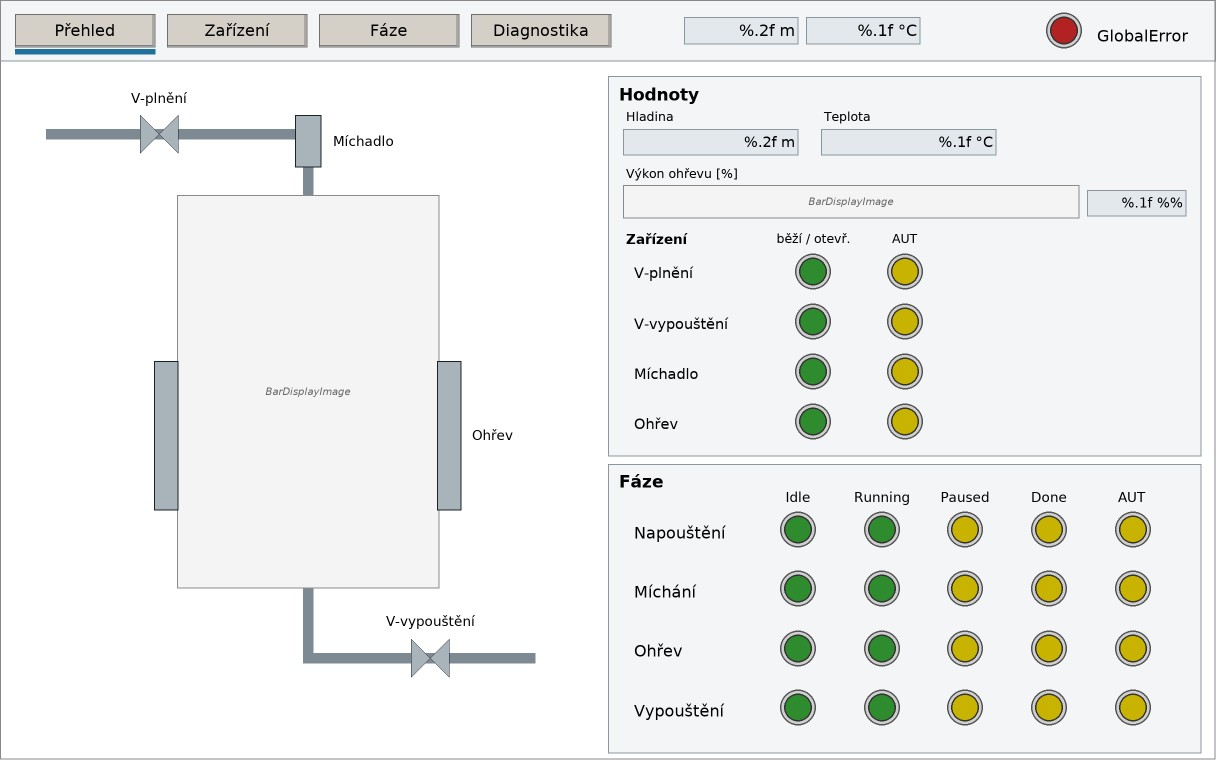
VISUALIZATION Prehled  // 1216x760
    Rectangle (0,0 1216x61)
    Button (15,14 140x33), "Přehled"
        OnMouseClick: change screen: Prehled
    Rectangle (15,49 140x5)
    Button (167,14 140x33), "Zařízení"
        OnMouseClick: change screen: Zarizeni
    Button (319,14 140x33), "Fáze"
        OnMouseClick: change screen: Faze
    Button (471,14 140x33), "Diagnostika"
        OnMouseClick: change screen: Diagnostika
    Rectangle (684,17 114x27), "%.2f m", text variable: Global.Tank1.Filling.WaterLevel
    Rectangle (806,17 114x27), "%.1f °C", text variable: Global.Tank1.Heating.WaterTemp
    Lamp1 (1041,10 46x41), variable: Global.Tank1.GlobalError, style: Lamp-Lamp1-Red
    Label (1094,23 126x26), "GlobalError"
    Rectangle (46,129 267x10)
    Rectangle (303,129 10x68)
    Rectangle (303,586 10x77)
    Rectangle (303,653 232x10)
    BarDisplayImage (177,195 262x393), value: Global.Tank1.Filling.WaterLevel, style: BarDisplayImage-Gray, scale format: %.1f, scale 0..2
    Polygon (140,115) (178,153) (178,115) (140,153) (140,153), colour toggle: Global.Tank1.ValveFilling.State.Open
    Label (121,87 76x23), "V-plnění"
    Polygon (411,639) (449,677) (449,639) (411,677) (411,677), colour toggle: Global.Tank1.ValveDraining.State.Open
    Label (385,610 91x23), "V-vypouštění"
    Rectangle (295,115 26x52), colour toggle: Global.Tank1.Mixer.State.Run
    Label (330,130 80x23), "Míchadlo"
    Rectangle (154,361 24x149), colour toggle: Global.Tank1.Heater.State.EnableOut
    Rectangle (437,361 24x149), colour toggle: Global.Tank1.Heater.State.EnableOut
    Label (469,424 52x23), "Ohřev"
    Rectangle (608,76 593x380)
    Label (616,81 87x27), "Hodnoty"
    Label (623,106 66x21), "Hladina"
    Rectangle (623,129 175x26), "%.2f m", text variable: Global.Tank1.Filling.WaterLevel
    Label (821,106 66x21), "Teplota"
    Rectangle (821,129 175x26), "%.1f °C", text variable: Global.Tank1.Heating.WaterTemp
    Label (623,163 142x21), "Výkon ohřevu [%]"
    BarDisplayImage (623,185 456x33), value: Global.Tank1.Heater.State.HeatingOut, style: BarDisplayImage-Gray, scale format: %.1f, scale 0..100
    Rectangle (1087,190 99x26), "%.1f %%", text variable: Global.Tank1.Heater.State.HeatingOut
    Label (623,228 80x23), "Zařízení"
    Label (768,228 91x21), "běží / otevř."
    Label (859,228 91x21), "AUT"
    Label (631,261 84x24), "V-plnění"
    Lamp1 (790,251 46x41), variable: Global.Tank1.ValveFilling.State.Open, style: Lamp-Lamp1-Green
    Lamp1 (882,251 46x41), variable: Global.Tank1.ValveFilling.State.AutCtrl, style: Lamp-Lamp1-Yellow
    Label (631,312 123x24), "V-vypouštění"
    Lamp1 (790,301 46x41), variable: Global.Tank1.ValveDraining.State.Open, style: Lamp-Lamp1-Green
    Lamp1 (882,301 46x41), variable: Global.Tank1.ValveDraining.State.AutCtrl, style: Lamp-Lamp1-Yellow
    Label (631,362 84x24), "Míchadlo"
    Lamp1 (790,351 46x41), variable: Global.Tank1.Mixer.State.Run, style: Lamp-Lamp1-Green
    Lamp1 (882,351 46x41), variable: Global.Tank1.Mixer.State.AutCtrl, style: Lamp-Lamp1-Yellow
    Label (631,412 55x24), "Ohřev"
    Lamp1 (790,401 46x41), variable: Global.Tank1.Heater.State.EnableOut, style: Lamp-Lamp1-Green
    Lamp1 (882,401 46x41), variable: Global.Tank1.Heater.State.AutCtrl, style: Lamp-Lamp1-Yellow
    Rectangle (608,464 593x289)
    Label (616,468 53x27), "Fáze"
    Label (760,486 76x23), "Idle"
    Label (844,486 76x23), "Running"
    Label (927,486 76x23), "Paused"
    Label (1011,486 76x23), "Done"
    Label (1094,486 76x23), "AUT"
    Label (631,520 116x26), "Napouštění"
    Lamp1 (775,509 46x41), variable: Global.Tank1.Filling.State.Idle, style: Lamp-Lamp1-Green
    Lamp1 (859,509 46x41), variable: Global.Tank1.Filling.State.Running, style: Lamp-Lamp1-Green
    Lamp1 (942,509 46x41), variable: Global.Tank1.Filling.State.Paused, style: Lamp-Lamp1-Yellow
    Lamp1 (1026,509 46x41), variable: Global.Tank1.Filling.State.Done, style: Lamp-Lamp1-Yellow
    Lamp1 (1110,509 46x41), variable: Global.Tank1.Filling.State.AutCtrl, style: Lamp-Lamp1-Yellow
    Label (631,579 83x26), "Míchání"
    Lamp1 (775,568 46x41), variable: Global.Tank1.Mixing.State.Idle, style: Lamp-Lamp1-Green
    Lamp1 (859,568 46x41), variable: Global.Tank1.Mixing.State.Running, style: Lamp-Lamp1-Green
    Lamp1 (942,568 46x41), variable: Global.Tank1.Mixing.State.Paused, style: Lamp-Lamp1-Yellow
    Lamp1 (1026,568 46x41), variable: Global.Tank1.Mixing.State.Done, style: Lamp-Lamp1-Yellow
    Lamp1 (1110,568 46x41), variable: Global.Tank1.Mixing.State.AutCtrl, style: Lamp-Lamp1-Yellow
    Label (631,638 62x26), "Ohřev"
    Lamp1 (775,628 46x41), variable: Global.Tank1.Heating.State.Idle, style: Lamp-Lamp1-Green
    Lamp1 (859,628 46x41), variable: Global.Tank1.Heating.State.Running, style: Lamp-Lamp1-Green
    Lamp1 (942,628 46x41), variable: Global.Tank1.Heating.State.Paused, style: Lamp-Lamp1-Yellow
    Lamp1 (1026,628 46x41), variable: Global.Tank1.Heating.State.Done, style: Lamp-Lamp1-Yellow
    Lamp1 (1110,628 46x41), variable: Global.Tank1.Heating.State.AutCtrl, style: Lamp-Lamp1-Yellow
    Label (631,698 116x26), "Vypouštění"
    Lamp1 (775,687 46x41), variable: Global.Tank1.Draining.State.Idle, style: Lamp-Lamp1-Green
    Lamp1 (859,687 46x41), variable: Global.Tank1.Draining.State.Running, style: Lamp-Lamp1-Green
    Lamp1 (942,687 46x41), variable: Global.Tank1.Draining.State.Paused, style: Lamp-Lamp1-Yellow
    Lamp1 (1026,687 46x41), variable: Global.Tank1.Draining.State.Done, style: Lamp-Lamp1-Yellow
    Lamp1 (1110,687 46x41), variable: Global.Tank1.Draining.State.AutCtrl, style: Lamp-Lamp1-Yellow
END_VISUALIZATION

// ---- VISUs/Zarizeni.TcVIS
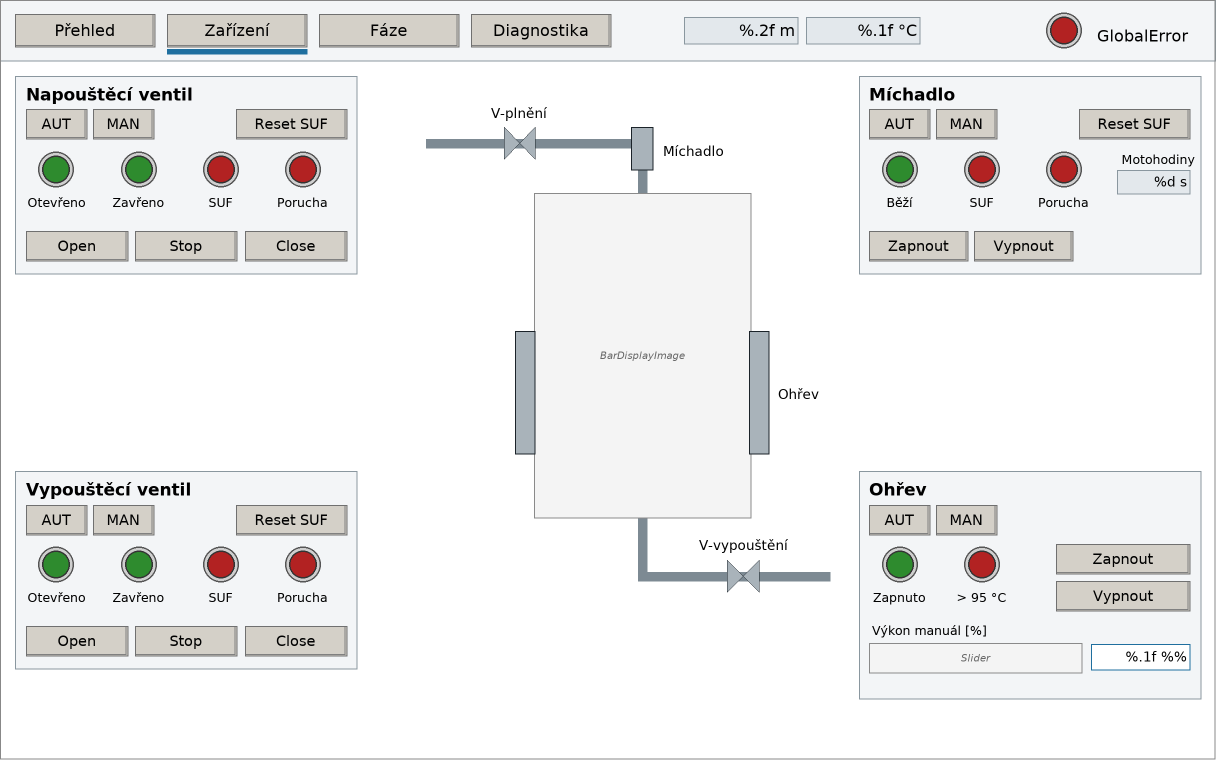
VISUALIZATION Zarizeni  // 1216x760
    Rectangle (0,0 1216x61)
    Button (15,14 140x33), "Přehled"
        OnMouseClick: change screen: Prehled
    Button (167,14 140x33), "Zařízení"
        OnMouseClick: change screen: Zarizeni
    Rectangle (167,49 140x5)
    Button (319,14 140x33), "Fáze"
        OnMouseClick: change screen: Faze
    Button (471,14 140x33), "Diagnostika"
        OnMouseClick: change screen: Diagnostika
    Rectangle (684,17 114x27), "%.2f m", text variable: Global.Tank1.Filling.WaterLevel
    Rectangle (806,17 114x27), "%.1f °C", text variable: Global.Tank1.Heating.WaterTemp
    Lamp1 (1041,10 46x41), variable: Global.Tank1.GlobalError, style: Lamp-Lamp1-Red
    Label (1094,23 126x26), "GlobalError"
    Rectangle (426,139 221x9)
    Rectangle (638,139 9x56)
    Rectangle (638,517 9x64)
    Rectangle (638,572 192x9)
    BarDisplayImage (534,193 217x325), value: Global.Tank1.Filling.WaterLevel, style: BarDisplayImage-Gray, scale format: %.1f, scale 0..2
    Polygon (504,127) (535,159) (535,127) (504,159) (504,159), colour toggle: Global.Tank1.ValveFilling.State.Open
    Label (481,102 76x23), "V-plnění"
    Polygon (727,560) (759,592) (759,560) (727,592) (727,592), colour toggle: Global.Tank1.ValveDraining.State.Open
    Label (698,534 91x23), "V-vypouštění"
    Rectangle (631,127 22x43), colour toggle: Global.Tank1.Mixer.State.Run
    Label (660,140 80x23), "Míchadlo"
    Rectangle (515,331 20x123), colour toggle: Global.Tank1.Heater.State.EnableOut
    Rectangle (749,331 20x123), colour toggle: Global.Tank1.Heater.State.EnableOut
    Label (775,383 52x23), "Ohřev"
    Rectangle (15,76 342x198)
    Label (23,81 201x27), "Napouštěcí ventil"
    Button (26,109 61x30), "AUT", colour toggle: Global.Tank1.ValveFilling.State.AutCtrl
        tap Global.Tank1.ValveFilling.Cmd.AutCtrl
    Button (93,109 61x30), "MAN", colour toggle: Global.Tank1.ValveFilling.State.ManCtrl
        tap Global.Tank1.ValveFilling.Cmd.ManCtrl
    Button (236,109 111x30), "Reset SUF", colour toggle: Global.Tank1.ValveFilling.State.StartupFail
        tap Global.Tank1.ValveFilling.Cmd.ResetSUF
    Lamp1 (33,149 46x41), variable: Global.Tank1.ValveFilling.State.Open, style: Lamp-Lamp1-Green
    Label (11,192 91x21), "Otevřeno"
    Lamp1 (116,149 46x41), variable: Global.Tank1.ValveFilling.State.Closed, style: Lamp-Lamp1-Green
    Label (93,192 91x21), "Zavřeno"
    Lamp1 (198,149 46x41), variable: Global.Tank1.ValveFilling.State.StartupFail, style: Lamp-Lamp1-Red
    Label (175,192 91x21), "SUF"
    Lamp1 (280,149 46x41), variable: Global.Tank1.ValveFilling.State.Err, style: Lamp-Lamp1-Red
    Label (257,192 91x21), "Porucha"
    Button (26,231 102x30), "Open", colour toggle: Global.Tank1.ValveFilling.State.Open
        tap Global.Tank1.ValveFilling.Cmd.OpenMan
    Button (135,231 102x30), "Stop"
        tap Global.Tank1.ValveFilling.Cmd.StopMan
    Button (245,231 102x30), "Close", colour toggle: Global.Tank1.ValveFilling.State.Closed
        tap Global.Tank1.ValveFilling.Cmd.CloseMan
    Rectangle (859,76 342x198)
    Label (866,81 99x27), "Míchadlo"
    Button (869,109 61x30), "AUT", colour toggle: Global.Tank1.Mixer.State.AutCtrl
        tap Global.Tank1.Mixer.Cmd.AutCtrl
    Button (936,109 61x30), "MAN", colour toggle: Global.Tank1.Mixer.State.ManCtrl
        tap Global.Tank1.Mixer.Cmd.ManCtrl
    Button (1079,109 111x30), "Reset SUF", colour toggle: Global.Tank1.Mixer.State.StartUpFail
        tap Global.Tank1.Mixer.Cmd.ResetSUF
    Lamp1 (877,149 46x41), variable: Global.Tank1.Mixer.State.Run, style: Lamp-Lamp1-Green
    Label (854,192 91x21), "Běží"
    Lamp1 (959,149 46x41), variable: Global.Tank1.Mixer.State.StartUpFail, style: Lamp-Lamp1-Red
    Label (936,192 91x21), "SUF"
    Lamp1 (1041,149 46x41), variable: Global.Tank1.Mixer.State.Err, style: Lamp-Lamp1-Red
    Label (1018,192 91x21), "Porucha"
    Button (869,231 99x30), "Zapnout", colour toggle: Global.Tank1.Mixer.State.Run
        tap Global.Tank1.Mixer.Cmd.TurnOnMan
    Button (974,231 99x30), "Vypnout"
        tap Global.Tank1.Mixer.Cmd.TurnOffMan
    Label (1122,149 73x21), "Motohodiny"
    Rectangle (1117,170 73x24), "%d s", text variable: Global.Tank1.Mixer.State.RT
    Rectangle (15,471 342x198)
    Label (23,476 201x27), "Vypouštěcí ventil"
    Button (26,505 61x30), "AUT", colour toggle: Global.Tank1.ValveDraining.State.AutCtrl
        tap Global.Tank1.ValveDraining.Cmd.AutCtrl
    Button (93,505 61x30), "MAN", colour toggle: Global.Tank1.ValveDraining.State.ManCtrl
        tap Global.Tank1.ValveDraining.Cmd.ManCtrl
    Button (236,505 111x30), "Reset SUF", colour toggle: Global.Tank1.ValveDraining.State.StartupFail
        tap Global.Tank1.ValveDraining.Cmd.ResetSUF
    Lamp1 (33,544 46x41), variable: Global.Tank1.ValveDraining.State.Open, style: Lamp-Lamp1-Green
    Label (11,587 91x21), "Otevřeno"
    Lamp1 (116,544 46x41), variable: Global.Tank1.ValveDraining.State.Closed, style: Lamp-Lamp1-Green
    Label (93,587 91x21), "Zavřeno"
    Lamp1 (198,544 46x41), variable: Global.Tank1.ValveDraining.State.StartupFail, style: Lamp-Lamp1-Red
    Label (175,587 91x21), "SUF"
    Lamp1 (280,544 46x41), variable: Global.Tank1.ValveDraining.State.Err, style: Lamp-Lamp1-Red
    Label (257,587 91x21), "Porucha"
    Button (26,626 102x30), "Open", colour toggle: Global.Tank1.ValveDraining.State.Open
        tap Global.Tank1.ValveDraining.Cmd.OpenMan
    Button (135,626 102x30), "Stop"
        tap Global.Tank1.ValveDraining.Cmd.StopMan
    Button (245,626 102x30), "Close", colour toggle: Global.Tank1.ValveDraining.State.Closed
        tap Global.Tank1.ValveDraining.Cmd.CloseMan
    Rectangle (859,471 342x228)
    Label (866,476 65x27), "Ohřev"
    Button (869,505 61x30), "AUT", colour toggle: Global.Tank1.Heater.State.AutCtrl
        tap Global.Tank1.Heater.Cmd.AutCtrl
    Button (936,505 61x30), "MAN", colour toggle: Global.Tank1.Heater.State.ManCtrl
        tap Global.Tank1.Heater.Cmd.ManCtrl
    Lamp1 (877,544 46x41), variable: Global.Tank1.Heater.State.EnableOut, style: Lamp-Lamp1-Green
    Label (854,587 91x21), "Zapnuto"
    Lamp1 (959,544 46x41), variable: Global.Tank1.Heater.State.GenErr, style: Lamp-Lamp1-Red
    Label (936,587 91x21), "> 95 °C"
    Button (1056,544 134x30), "Zapnout", colour toggle: Global.Tank1.Heater.State.EnableOut
        tap Global.Tank1.Heater.Cmd.TurnOnMan
    Button (1056,581 134x30), "Vypnout"
        tap Global.Tank1.Heater.Cmd.TurnOffMan
    Label (869,620 142x21), "Výkon manuál [%]"
    Slider (869,643 213x30), variable: Global.Tank1.Heater.ParamHeatingPowerManual, scale 0..100
    Rectangle (1091,644 99x26), "%.1f %%", text variable: Global.Tank1.Heater.ParamHeatingPowerManual
        OnMouseClick: write the text variable via Default
END_VISUALIZATION
